(* IEC 61131-3 sources: daoli-st-library/DL_Process (part 29) *)

(* ---- FB_DL_ConveyorAccumGateSeq.st ---- *)
//==============================================================================
// 功能块：FB_DL_ConveyorAccumGateSeq ｜ 中文名称：输送线积放闸门三态序列编排
// 所属子库：DL_Process ｜ 版本：v1.0.0 ｜ 日期：2026-11-23
// 兼容：CODESYS V3.5+ / TwinCAT 3 / 汇川 InoProShop（纯 IEC 61131-3 第 3 版，零方言）
// 功能描述：积放/释放/满流三态编排：积放相闸门关闭、物料在积放位堆积；
//           积放位满且下游可收 → 释放相（闸门开，按 tKick 节拍向下游发
//           bDownKick 联动脉冲）；积放位满且下游不可收 → 满流相（闸门关 +
//           bUpstreamStop 请求上游节拍停止，信息级留痕）。闸门开启设最小
//           开门时长防阀/闸颤振；释放完成回积放或待机。下游节拍联动由
//           自复位周期窗 TON 生成（IN := NOT tonXxx.Q，R188 口径）。
// 开源溯源 (Origin)：原创实现（s9-conv 输送工程惯例深化，零外部源码行，
//           clean-room 独立编写）
// 公开接口清单：输入 bEn / bUpstreamRun / bFullSens / bDownReady /
//               tMinGate / tKick；
//               输出 bGateOpen / bUpstreamStop / bDownKick / eState /
//               uErrCode / bValid
// 单位表：tMinGate[ms] / tKick[ms]，其余 BOOL 引脚无量纲
// 输入契约：bFullSens 为积放位满传感，bDownReady 为下游可收声明，均经
//           IO 映射层注入；tMinGate 防闸门颤振下限；tKick 节拍周期。
// 输出契约：bGateOpen 请求级闸门开指令（执行器驱动须上层联锁）；
//           bDownKick 单拍节拍脉冲；uErrCode 信息级不锁存；
//           bValid 恒 TRUE（本件无故障级条件）。
// 错误码表：16#0005_3050 信息级（满流节拍停止请求激活，不置 bError）/
//           16#0005_3051 信息级（非法状态兜底入安全侧待机，不置 bError）/
//           16#0005_3052 预留禁用（不得挪用）
// 状态机：E_DL_AccumGateState（本文件唯一定义，全库唯一属主）：
//           eIdle = 0 / eAccumulating = 10 / eFullStop = 20 / eReleasing = 30
// 边界行为：① 闸门默认关（所有相默认值安全侧），开门仅释放相声明；
//           ② 最小开门时长未满不关门（防颤振）；
//           ③ 节拍脉冲 TON 自复位（IN := NOT tonKick.Q），每拍无条件刷新；
//           ④ 撤使能任意相回待机且闸门关（门控挂状态量）；
//           ⑤ CASE 带 ELSE 非法态兜底回 eIdle（信息级留痕）；
//           ⑥ 本件无故障级条件，不设 bError（码表与实现对齐，不虚声明）。
// 修订历史：v1.0.0 2026-11-23 首版（R73 派单 · 批 2 · 序 6）
//==============================================================================

(*------------------------------------------------------------------------------
 * 枚举: E_DL_AccumGateState（归属本功能块，同文件发布，全库唯一属主）
 * 含义: 积放闸门序列相位，成员与 CASE 标签双向完备。
 *-----------------------------------------------------------------------------*)
TYPE E_DL_AccumGateState :
(
    eIdle         := 0,   // 待机：闸门关，等使能与上游 / Idle, gate closed
    eAccumulating := 10,  // 积放中：闸门关，物料堆积 / Accumulating, gate closed, stock piling
    eFullStop     := 20,  // 满流：闸门关 + 上游节拍停止请求 / Full, gate closed and upstream stop requested
    eReleasing    := 30   // 释放中：闸门开 + 下游节拍联动脉冲 / Releasing, gate open with downstream kick pulses
);
END_TYPE

(*==============================================================================
 * 功能块: FB_DL_ConveyorAccumGateSeq
 * 调用约定: 每个扫描周期无条件调用一次；实例状态全部驻留于私有变量。
 * 调用示例: accumGate(bEn := bLineEn, bUpstreamRun := bConvUpRun,
 *                     bFullSens := bAccumFull, bDownReady := bDownCS,
 *                     tMinGate := T#2S, tKick := T#1S);
 *          bGateOpen 驱动闸门电磁阀（经输出映射层），bDownKick 作下游
 *          节拍联动脉冲接入下游段使能合取。
 * 组装说明: ① 闸门驱动输出须在上层输出映射层复加机械限位联锁，本件
 *             bGateOpen 属请求级信号（红线 R2：零物理地址）；
 *           ② bFullSens / bDownReady 传感引脚经 PRG_IoMapping 读入注入；
 *           ③ tKick 节拍脉冲为单拍有效量，上层沿检测可省（直接作使能
 *             窗合取），如需展宽请串 FB_DL_PulseStretch；
 *           ④ 多级积放串联时，本级 bDownReady 取下级 accumGate.bGateOpen
 *             的取反（下级开门期间本级视为不可收）。
 *==============================================================================*)
FUNCTION_BLOCK FB_DL_ConveyorAccumGateSeq
VAR_INPUT
    bEn          : BOOL := FALSE;     // 使能（FALSE 任意相回待机）/ Enable, FALSE returns to idle from any phase
    bUpstreamRun : BOOL := FALSE;     // 上游段运行中 / Upstream section running
    bFullSens    : BOOL := FALSE;     // 积放位满传感器 / Accumulation zone full sensor
    bDownReady   : BOOL := FALSE;     // 下游可接收声明 / Downstream ready to receive
    tMinGate     : TIME := T#2S;      // 最小开门时长 [ms]，防闸门颤振 / Minimum gate-open duration [ms], anti-chatter
    tKick        : TIME := T#1S;      // 下游节拍联动脉冲周期 [ms] / Downstream kick pulse period [ms]
END_VAR
VAR_OUTPUT
    bGateOpen    : BOOL;              // 闸门开指令（仅释放相）/ Gate open command, releasing phase only
    bUpstreamStop: BOOL;              // 上游节拍停止请求（满流相）/ Upstream stop request, full phase
    bDownKick    : BOOL;              // 下游节拍联动脉冲（单拍有效）/ Downstream kick pulse, single-scan
    eState       : E_DL_AccumGateState; // 序列当前相位 / Current sequence phase
    uErrCode     : UDINT;             // 信息级码，0 = 无信息 / Info-level code, 0 = none
    bValid       : BOOL;              // 输出可用标志 / Outputs usable flag
END_VAR
VAR
    tonMinGate   : TON;               // 最小开门时长定时器，每拍无条件刷新 / Minimum gate-open timer, refreshed every scan
    tonKick      : TON;               // 节拍脉冲自复位定时器，每拍无条件刷新 / Kick pulse self-reset timer, refreshed every scan
END_VAR
VAR CONSTANT
    DL_CG_CODE_FULL : UDINT := 16#0005_3050; // 信息级：满流停止请求码 / Info code: full-flow stop request
    DL_CG_CODE_ILL  : UDINT := 16#0005_3051; // 信息级：非法状态兜底码 / Info code: illegal state fallback
END_VAR

// ---- 段 1｜定时器无条件刷新（红线 R7：禁入条件分支；tonKick 自复位 R188）----
tonMinGate(IN := (eState = E_DL_AccumGateState.eReleasing), PT := tMinGate); // 开门计时按相断输入 / Gate timer input per phase
tonKick(IN := (eState = E_DL_AccumGateState.eReleasing)
        AND bDownReady AND NOT tonKick.Q, PT := tKick); // 周期窗自复位（R188 口径）/ Self-resetting window per R188

// ---- 段 2｜出口默认值：入口即赋安全侧确定值 ----
bGateOpen     := FALSE;             // 闸门默认关（安全侧）/ Gate preset closed, safe side
bUpstreamStop := FALSE;             // 上游停止请求默认 FALSE / Upstream stop preset FALSE
bDownKick     := FALSE;             // 节拍脉冲默认 FALSE（相内重映射）/ Kick pulse preset FALSE
uErrCode      := 16#0000_0000;      // 信息码每拍重算（信息级不锁存）/ Info code recomputed, never latched
bValid        := TRUE;              // 可用标志默认 TRUE / Usable flag preset TRUE

// ---- 段 3｜序列状态机（CASE 带 ELSE；满流先于释放判决防抢跑）----
CASE eState OF
    E_DL_AccumGateState.eIdle:        // 待机相：闸门关，等使能
        IF bEn AND bUpstreamRun THEN
            eState := E_DL_AccumGateState.eAccumulating; // 进入积放相 / Enter accumulating
        END_IF

    E_DL_AccumGateState.eAccumulating:// 积放相：闸门关，堆积至满
        IF NOT (bEn AND bUpstreamRun) THEN
            eState := E_DL_AccumGateState.eIdle; // 撤条件回待机 / Conditions lost, back to idle
        ELSIF bFullSens THEN
            IF bDownReady THEN        // 满且下游可收 → 释放（满流先判下游）/ Full and downstream ready, release first
                eState := E_DL_AccumGateState.eReleasing;
            ELSE                      // 满且下游不可收 → 满流停止请求 / Full and not ready, full-stop
                eState := E_DL_AccumGateState.eFullStop;
            END_IF
        END_IF

    E_DL_AccumGateState.eFullStop:    // 满流相：闸门关 + 上游停止请求（信息级）
        bUpstreamStop := TRUE;        // 上游节拍停止请求 / Upstream stop request
        uErrCode := DL_CG_CODE_FULL;  // 信息级留痕（每拍重算，不置 bError）/ Info trace, no fault flag
        IF bDownReady THEN            // 下游恢复可收 → 转释放 / Downstream ready, go release
            eState := E_DL_AccumGateState.eReleasing;
        ELSIF NOT bFullSens THEN      // 积放位已不满（上游停后消化）→ 回积放 / Zone drained, back to accumulating
            eState := E_DL_AccumGateState.eAccumulating;
        END_IF

    E_DL_AccumGateState.eReleasing:   // 释放相：闸门开 + 节拍联动脉冲
        bGateOpen := TRUE;            // 闸门开声明 / Gate open declared
        bDownKick := tonKick.Q AND bDownReady; // 节拍联动脉冲（单拍有效）/ Kick pulse, single-scan
        IF NOT bEn THEN
            eState := E_DL_AccumGateState.eIdle; // 撤使能回待机 / Disable, back to idle
        ELSIF tonMinGate.Q AND (NOT bFullSens) THEN
            IF bUpstreamRun THEN
                eState := E_DL_AccumGateState.eAccumulating; // 释放完回积放 / Done, back to accumulating
            ELSE
                eState := E_DL_AccumGateState.eIdle; // 释放完且上游停回待机 / Done and upstream stopped, back to idle
            END_IF
        ELSIF (NOT bDownReady) AND tonMinGate.Q THEN
            eState := E_DL_AccumGateState.eFullStop; // 下游中途不可收 → 满流 / Downstream lost, go full-stop
        END_IF

    ELSE                              // 非法状态兜底（R21：CASE 必带 ELSE）
        eState   := E_DL_AccumGateState.eIdle; // 拦截非法值回待机（安全侧闸门关）/ Catch illegal value to idle, gate closed
        uErrCode := DL_CG_CODE_ILL;   // 信息级兜底留痕（不置 bError）/ Info-level fallback trace
END_CASE

// ---- 段 4｜统一出口：撤使能兜底（门控挂状态量）----
IF NOT bEn THEN
    IF eState <> E_DL_AccumGateState.eIdle THEN
        eState := E_DL_AccumGateState.eIdle; // 回待机 / Back to idle
    END_IF
    bGateOpen := FALSE;               // 闸门强制关 / Gate forced closed
    bUpstreamStop := FALSE;           // 停止请求撤除 / Stop request withdrawn
END_IF
END_FUNCTION_BLOCK

(* ---- FB_DL_ConveyorDirMismatch.st ---- *)
(*
  FB_DL_ConveyorDirMismatch  —  输送线停机方向失配独立诊断窗（反窜/倒滑） / Conveyor stopped-state direction mismatch diagnostic window
  分类 Category : DL_Process
  版本 Version  : 1.0.1
  来源 Source   : t2-7-packml — 终审立项独立诊断增强（复用 FB_DL_ConveyorZone 光电语义）
  溯源 Origin   : clean-room 实现，未复制任何源码行
  功能 Function : 1) 停机判据用当拍量（NOT bMotorRun）；停机后经 tSettle 静置窗进 eWatch
                  监视相，独立诊断窗 TON（tonDiagBack/tonDiagSlide）与运行窗分实例；
                  2) 反窜诊断：停机监视相中入口光电持续遮挡（电平承载）超 tDiagWin
                  → 故障级 036D 独立锁存（R190 归因唯一）；
                  3) 倒滑诊断：停机监视相中出口光电持续遮挡超 tDiagWin
                  → 故障级 036E 独立锁存；
                  4) 相位机 CASE 全覆盖 + ELSE 兜底落 036F；诊断窗 TON 无条件
                  周期刷新且 IN 用光电电平承载（门控沿与计时基解耦，与
                  FB_DL_ConveyorZone run-on 语义分工：那件管运行清区，本件管停机反常）。
  返修记录 Rework  :
    2026-11-19  v1.0.1  R42 P0-1 严重返修：v1.0.0 诊断窗 TON 的 IN 由光电沿实例
                        rtPeEntry.Q/rtPeDis.Q（单拍量）门控——沿为单拍脉冲，TON 计时基
                        下一拍即断，结构性永不到时（P0 派单缺陷①）。修复要点：TON 的 IN
                        改由光电电平（bPEEntry/bPEDischarge）与监视相单相等式承载，
                        沿实例随结构性缺陷一并移除；对外接口签名不变；
                        光电语义改为「持续遮挡超 tDiagWin」判反窜/倒滑。
  边界 Boundary : ① 运行恢复（bMotorRun 当拍 TRUE）即回 eIdle，诊断窗自动清；
                  ② 解除式全当拍量（R240 落地）：rtReset.Q AND NOT bMotorRun，逐 BOOL 标注见段 4；
                  ③ 组态闸：tSettle/tDiagWin <= 0 → 036F 同级锁存（组态与兜底归并声明于码表）；
                  ④ 无 GVL 依赖：纯引脚输入输出，无外部变量引用，无物理 IO 地址。
  依赖 Depends  : 与 FB_DL_ConveyorZone 光电/run-on 语义分工对齐（不实例化）；Standard.library（TON / R_TRIG / F_TRIG）
  码表 Error codes（Process 段 0005，窗口 036D~036F / 0495~0497）:
    16#0005_036D 故障级：反窜检出锁存（停机监视相入口光电持续遮挡超 tDiagWin），锁存至 bReset
    16#0005_036E 故障级：倒滑检出锁存（停机监视相出口光电持续遮挡超 tDiagWin），锁存至 bReset
    16#0005_036F 故障级：相位落 ELSE 兜底或组态非法（静置/诊断窗域非法），锁存至 bReset
    16#0005_0495 信息级：诊断窗激活沿（进入 eWatch）
    16#0005_0496 信息级：反窜解除沿（复位清锁存）
    16#0005_0497 信息级：倒滑解除沿（复位清锁存）
  修订历史 Revision :
    2026-11-19  v1.0.0  R41 首版（批次 4 · 序号 5）
    2026-11-19  v1.0.1  R42 P0-1 严重返修（见返修记录节）
*)

TYPE E_DL_CdmState :
(
    eIdle   := 0,    // 空闲：运行中或无停机事件 / Idle, running or no stop event
    eSettle := 10,   // 静置：停机确认窗 / Settle, stopped confirm window
    eWatch  := 20,   // 监视：独立诊断窗开启 / Watch, diagnostic window open
    eFault  := 90    // 故障：反窜或倒滑锁定 / Fault, latched
);
END_TYPE

FUNCTION_BLOCK FB_DL_ConveyorDirMismatch
VAR_INPUT
    bMotorRun    : BOOL := FALSE;     // 驱动运行反馈，TRUE = 运行中 [-] / Drive running feedback
    bFwdCmd      : BOOL := TRUE;      // 运行方向指令，TRUE = 正向（诊断口径记录用）[-] / Direction command
    bPEEntry     : BOOL := FALSE;     // 入口光电，TRUE = 遮挡 [-] / Entry photoeye, TRUE = blocked
    bPEDischarge : BOOL := FALSE;     // 出口光电，TRUE = 遮挡 [-] / Discharge photoeye, TRUE = blocked
    tSettle      : TIME := T#2S;      // 停机静置窗 [ms]，域 > 0 / Stop settle window
    tDiagWin     : TIME := T#5S;      // 独立诊断窗 [ms]，域 > 0 / Diagnostic window
    bReset       : BOOL := FALSE;     // 复位，上升沿清故障锁存 / Reset edge clears fault latch
END_VAR
VAR_OUTPUT
    eState       : E_DL_CdmState;     // 状态出口，段尾单点映射 / State outlet
    bBackFlow    : BOOL;              // 反窜独立锁存出口 [-] / Back-flow latch outlet
    bSlideBack   : BOOL;              // 倒滑独立锁存出口 [-] / Slide-back latch outlet
    bFault       : BOOL;              // 聚合故障标志 / Aggregate fault flag
    bError       : BOOL;              // 故障级标志（与聚合锁存同源）/ Fault flag
    nErrId       : UDINT;             // 事件码，0 = 无事件 / Event code
END_VAR
VAR
    tonSettle    : TON;               // 停机静置窗 TON（与运行窗分实例），无条件刷新 / Settle timer
    tonDiagBack  : TON;               // 反窜独立诊断窗 TON，无条件刷新 / Back-flow diagnostic timer
    tonDiagSlide : TON;               // 倒滑独立诊断窗 TON，无条件刷新 / Slide-back diagnostic timer
    rtPeEntry    : R_TRIG;            // 入口光电沿实例（v1.0.1 已移除判据用途，保留供上层诊断镜像）；
                                       // 上层不引用时可在组装层删除 / Entry photoeye edge instance (no longer gating)
    rtPeDis      : R_TRIG;            // 出口光电沿实例（v1.0.1 已移除判据用途，前述解除判据）/ Discharge photoeye edge instance
    rtReset      : R_TRIG;            // 复位沿实例，无条件刷新 / Reset edge instance
    _eState      : E_DL_CdmState := E_DL_CdmState.eIdle;  // 内部相位（CASE 唯一写入目标）/ Internal phase
    _bStopped    : BOOL;              // 停机当拍量 [-] / Stopped current-scan flag
    _bBackLat    : BOOL;              // 反窜锁存位（锁存量）/ Back-flow latch bit
    _bSlideLat   : BOOL;              // 倒滑锁存位（锁存量）/ Slide-back latch bit
    _bCfgBad     : BOOL;              // 组态锁存位（锁存量）/ Config-fault latch bit
    _uFault      : UDINT;             // 故障码锁存（锁存量）/ Latched fault code
    _uInfo       : UDINT;             // 信息码，每拍重算 / Transient info code
    _bWatchPrev  : BOOL;              // 上拍监视相镜像（激活沿判据）/ Previous watch mirror
    _bBackOkPrev : BOOL;              // 上拍反窜无锁存镜像（解除沿判据）/ Previous back-clear mirror
    _bSlideOkPrev: BOOL;              // 上拍倒滑无锁存镜像（解除沿判据）/ Previous slide-clear mirror
END_VAR

(* —— 段 0：定时器与沿实例无条件周期刷新（禁置于 IF/CASE 内） —— *)
_bStopped := NOT bMotorRun;                          // 停机判据（当拍量）
rtPeEntry(CLK := bPEEntry);                          // 入口光电沿（每拍必调）
rtPeDis(CLK := bPEDischarge);                        // 出口光电沿（每拍必调）
rtReset(CLK := bReset);                              // 复位沿（每拍必调）
tonSettle(IN := (_eState = E_DL_CdmState.eSettle), PT := tSettle);              // 静置窗（单相独占）
tonDiagBack(IN := (_eState = E_DL_CdmState.eWatch) AND bPEEntry, PT := tDiagWin);
                                                     // 反窜诊断窗（光电电平承载，门控沿与计时基解耦，每拍必调）
tonDiagSlide(IN := (_eState = E_DL_CdmState.eWatch) AND bPEDischarge, PT := tDiagWin);
                                                     // 倒滑诊断窗（光电电平承载，前述解除判据，每拍必调）

(* —— 段 1：单拍量预清零（锁存量 _uFault/_bBackLat/_bSlideLat/_bCfgBad 不入清单，禁同拍抹除） —— *)
_uInfo := 16#0000_0000;             // 信息码每拍重算
nErrId := 16#0000_0000;             // 事件码缺省无事件

(* —— 段 2：复位沿 + 组态域闸（当拍量判据） —— *)
IF rtReset.Q THEN                   // rtReset.Q = 当拍量
    _bBackLat := FALSE;             // 清反窜锁存位
    _bSlideLat := FALSE;            // 清倒滑锁存位
    _bCfgBad := FALSE;              // 清组态锁存位
    _uFault := 16#0000_0000;        // 清故障锁存码
END_IF
IF (TIME_TO_DINT(tSettle) <= 0) OR (TIME_TO_DINT(tDiagWin) <= 0) THEN
    _uFault := 16#0005_036F;        // 故障级：组态非法（归并兜底码，头注释③）
    _bCfgBad := TRUE;
END_IF

(* —— 段 3：双判据独立锁存（R190：反窜/倒滑归因唯一，各走独立码位与出口） —— *)
IF (_eState = E_DL_CdmState.eWatch) AND (NOT _bCfgBad) THEN
    IF tonDiagBack.Q THEN
        _uFault := 16#0005_036D;    // 故障级：反窜锁存
        _bBackLat := TRUE;
        _eState := E_DL_CdmState.eFault;
    ELSIF tonDiagSlide.Q THEN
        _uFault := 16#0005_036E;    // 故障级：倒滑锁存
        _bSlideLat := TRUE;
        _eState := E_DL_CdmState.eFault;
    END_IF
END_IF

(* —— 段 4：故障解除式（R240 落地，逐 BOOL 标注）：
     rtReset.Q = 当拍量；NOT bMotorRun = 当拍量；均不含锁存量（_bBackLat/_bSlideLat），
     解除边真实可达（复位沿在任意停机/运行拍均可到达）。 —— *)
IF rtReset.Q AND (NOT _bCfgBad) THEN
    IF _bBackLat THEN
        _uInfo := 16#0005_0496;     // 信息级：反窜解除沿
    END_IF
    IF _bSlideLat THEN
        _uInfo := 16#0005_0497;     // 信息级：倒滑解除沿（覆盖反窜解除沿，后到优先）
    END_IF
    _bBackLat := FALSE;             // 清反窜锁存位（锁存量，仅此当拍量解除沿可清）
    _bSlideLat := FALSE;            // 清倒滑锁存位（锁存量，仅解除沿可清）
    _uFault := 16#0000_0000;        // 清故障锁存码（锁存量，仅本当拍量解除沿可清）
END_IF

(* —— 段 5：相位机（CASE 全覆盖 + ELSE 兜底） —— *)
CASE _eState OF

E_DL_CdmState.eIdle:
    IF _bStopped AND (NOT _bCfgBad) THEN
        _eState := E_DL_CdmState.eSettle;   // 停机当拍：进静置相
    END_IF

E_DL_CdmState.eSettle:
    IF bMotorRun THEN                   // 运行恢复（当拍量）：回空闲
        _eState := E_DL_CdmState.eIdle;
    ELSIF tonSettle.Q THEN
        _uInfo := 16#0005_0495;         // 信息级：诊断窗激活沿
        _eState := E_DL_CdmState.eWatch;    // 静置通过：进监视相
    END_IF

E_DL_CdmState.eWatch:
    IF bMotorRun THEN                   // 运行恢复（当拍量）：回空闲（诊断窗自动清）
        _eState := E_DL_CdmState.eIdle;
    END_IF
    (* 反窜/倒滑检出与迁出在段 3 承载（独立诊断窗判据） *)

E_DL_CdmState.eFault:
    ;                                   // 故障相：等复位沿（段 4 承载迁出）

ELSE
    _uFault := 16#0005_036F;            // 故障级：非法相位兜底
    _bCfgBad := TRUE;
    _eState := E_DL_CdmState.eFault;    // 强制回故障相

END_CASE

(* —— 段 6：出口单点映射（名实同源；锁存码回放，禁同拍抹除） —— *)
bBackFlow := _bBackLat OR _bCfgBad;     // 反窜独立出口（组态坏并入安全侧）
bSlideBack := _bSlideLat OR _bCfgBad;   // 倒滑独立出口（前述解除判据）
bFault := _bBackLat OR _bSlideLat OR _bCfgBad;  // 聚合故障
IF bFault THEN
    nErrId := _uFault;              // 故障锁存码回放
ELSE
    nErrId := _uInfo;               // 信息码
END_IF
bError := bFault;                   // 故障标志与聚合锁存同源
eState := _eState;                  // 状态出口单点映射
_bWatchPrev := (_eState = E_DL_CdmState.eWatch);    // 激活沿判据快照
_bBackOkPrev := NOT _bBackLat;      // 解除沿判据快照
_bSlideOkPrev := NOT _bSlideLat;    // 解除沿判据快照

END_FUNCTION_BLOCK

(* ---- FB_DL_ConveyorMetalDetect.st ---- *)
// =====================================================================
// FB_DL_ConveyorMetalDetect.st
// 金属检测机剔除联动与过检率统计（延时排队/冻结补偿/确认超时锁存）
// Metal detector reject linkage and statistics FB
// 码位: 16#0005_0462 ~ 16#0005_0466 (本件独占 5 槽)
// 修改记录: R29 初版 (按 DISPATCH_R29 序 20)
// =====================================================================
FUNCTION_BLOCK FB_DL_ConveyorMetalDetect
VAR_INPUT
    bEnable        : BOOL  := FALSE;   // 使能 / Enable
    bReset         : BOOL  := FALSE;   // 复位（清统计）/ Reset
    bDetect        : BOOL  := FALSE;   // 检出脉冲（上升沿计数）/ Metal detected
    bRejectAck     : BOOL  := FALSE;   // 剔除完成确认 / Reject acknowledged
    fLineSpeed_mpm : REAL  := 0.0;     // 线速 0~200 m/min / Line speed [m/min]
    fSpeedMin_mpm  : REAL  := 1.0;     // 有效输送最小线速 >0 m/min / Min line speed [m/min]
    tRejectDelay   : TIME  := T#300MS; // 检测到剔除延时 T#10MS~T#5S / Reject delay [s]
    tRejectWidth   : TIME  := T#200MS; // 剔除脉冲宽度 T#20MS~T#2S / Reject pulse width [s]
    tAckMax        : TIME  := T#2S;    // 确认超时 T#100MS~T#30S / Ack timeout [s]
    uJamCnt        : USINT  := 3;      // 连续失败判卡滞次数 1~20 / Jam count
END_VAR
VAR_OUTPUT
    bRejectCmd     : BOOL;             // 剔除输出 / Reject command
    uDetectCnt     : UDINT;            // 累计检出数 / Detect count
    uRejectCnt     : UDINT;            // 累计已剔除数 / Rejected count
    fAckFailPct    : REAL;             // 确认失败率 0~100 % / Ack failure rate [%]
    bPending       : BOOL;             // 有剔除排队中 / Queue pending
    eErr           : UDINT;            // 错误码 / Error code
END_VAR
VAR
    rtrigDetect    : R_TRIG;           // 检出沿检测（无条件刷新）/ Detect edge detector
    tonDelay       : TON;              // 延时计时（皮带停时 IN 置 FALSE 冻结）/ Delay timer, frozen when belt stopped
    tonWidth       : TON;              // 脉宽计时 / Pulse width timer
    tonAck         : TON;              // 确认超时计时 / Ack timeout timer
    tDelayS        : REAL;             // 延时秒值 / Delay seconds [s]
    tWidthS        : REAL;             // 脉宽秒值 / Width seconds [s]
    tAckMaxS       : REAL;             // 超时秒值 / Timeout seconds [s]
    bDelaying      : BOOL;             // 延时排队中 / Delaying flag
    bRejecting     : BOOL;             // 剔除脉冲中 / Rejecting flag
    bAwaitingAck   : BOOL;             // 等确认中 / Awaiting ack flag
    bAckTimeoutLatch : BOOL := FALSE;  // 确认超时锁存 / Ack timeout latch
    uAckFailRun    : USINT;            // 连续确认失败计数 / Consecutive ack failure count
    bBeltMoving    : BOOL;             // 皮带运行判 / Belt moving flag
    uQueueDepth    : USINT;            // 排队深度（上限 8）/ Queue depth, cap 8
    xFirstScan     : BOOL  := TRUE;    // 首扫标记 / First-scan flag
END_VAR

// ---------------------------------------------------------------------
// 代码位表（本件独占，勿复用）:
//   16#0005_0462 信息 正常（无检出 / 剔除正常）
//   16#0005_0463 故障 线速非有限 / 任一 TIME 参数为 0 或非法
//   16#0005_0464 故障 fSpeedMin_mpm ≤ 0 / tRejectWidth ≥ tAckMax（组态错）
//   16#0005_0465 信息 排队冻结（fLineSpeed_mpm < fSpeedMin_mpm）→ 延时计时不走、bPending=TRUE
//   16#0005_0466 故障 单次确认超 tAckMax 或连续 uJamCnt 次失败 → 锁存；排队超 8 丢弃新检出同槽
// ---------------------------------------------------------------------

// ---- 时间转秒 / Times to seconds ----
tDelayS  := TIME_TO_REAL(tRejectDelay) / 1000.0;    // 延时秒 / Delay [s]
tWidthS  := TIME_TO_REAL(tRejectWidth) / 1000.0;    // 脉宽秒 / Width [s]
tAckMaxS := TIME_TO_REAL(tAckMax) / 1000.0;         // 超时秒 / Timeout [s]

// ---- 检出沿检测（无条件刷新）/ Detect edge, unconditional ----
rtrigDetect(CLK := bDetect);    // 沿检测 / Edge detection

// ---- 非有限与时间参数闸 / Finite and time validity gate ----
IF (fLineSpeed_mpm <> fLineSpeed_mpm) OR (ABS(fLineSpeed_mpm) >= 1.0E12)
   OR (fSpeedMin_mpm <> fSpeedMin_mpm) OR (ABS(fSpeedMin_mpm) >= 1.0E12)
   OR (tRejectDelay = T#0MS) OR (tDelayS < 0.01) OR (tDelayS > 5.0)
   OR (tRejectWidth = T#0MS) OR (tWidthS < 0.02) OR (tWidthS > 2.0)
   OR (tAckMax = T#0MS) OR (tAckMaxS < 0.1) OR (tAckMaxS > 30.0) THEN
    bRejectCmd := FALSE;        // 剔除撤销（安全侧）/ Reject off
    eErr := 16#0005_0463;       // 故障码 / Fault code
    RETURN;                     // 本拍结束 / End of cycle
END_IF

// ---- 组态错闸 / Configuration fault gate ----
IF (fSpeedMin_mpm <= 0.0) OR (tRejectWidth >= tAckMax) THEN
    bRejectCmd := FALSE;        // 剔除撤销 / Reject off
    eErr := 16#0005_0464;       // 故障码 / Fault code
    RETURN;                     // 本拍结束 / End of cycle
END_IF

// ---- 首扫初始化（R16 首扫纪律）/ First-scan initialization ----
IF xFirstScan THEN
    bRejectCmd := FALSE;        // 剔除初始关 / Reject init off
    bPending := FALSE;          // 排队复位 / Pending reset
    xFirstScan := FALSE;        // 清标记 / Clear flag
END_IF

// ---- 复位：清统计与队列 / Reset: clear statistics and queue ----
IF bReset THEN
    uDetectCnt := 0;            // 检出清零 / Detect cleared
    uRejectCnt := 0;            // 剔除清零 / Reject cleared
    fAckFailPct := 0.0;         // 失败率清零 / Fail rate cleared
    uAckFailRun := 0;           // 连败计数清零 / Fail run cleared
    bAckTimeoutLatch := FALSE;  // 锁存解除 / Latch released
    bDelaying := FALSE;         // 排队清空 / Queue cleared
    bRejecting := FALSE;        // 脉冲复位 / Pulse reset
    bAwaitingAck := FALSE;      // 等待复位 / Awaiting reset
    uQueueDepth := 0;           // 深度清零 / Depth cleared
END_IF

// ---- 使能撤销 / Disable ----
IF NOT bEnable THEN
    bRejectCmd := FALSE;        // 剔除撤销 / Reject off
    bDelaying := FALSE;         // 排队清空 / Queue cleared
    bRejecting := FALSE;        // 脉冲复位 / Pulse reset
    bAwaitingAck := FALSE;      // 等待复位 / Awaiting reset
    bPending := FALSE;          // 排队复位 / Pending reset
    eErr := 16#0005_0462;       // 信息级：空闲 / Info: idle
    RETURN;                     // 本拍结束 / End of cycle
END_IF

// ---- 确认超时锁存路径（漏剔是质量事故，宁可停线）/ Ack timeout latch path ----
IF bAckTimeoutLatch THEN
    bRejectCmd := FALSE;        // 剔除撤销 / Reject off
    eErr := 16#0005_0466;       // 故障码回放 / Fault code replay
    RETURN;                     // 本拍结束 / End of cycle
END_IF

// ---- 皮带运行判 / Belt moving check ----
bBeltMoving := (fLineSpeed_mpm >= fSpeedMin_mpm);   // 运行判 / Moving flag

// ---- 检出沿计数与排队（队列上限 8：超限丢弃并置槽 5，宁停线不漏剔）
// Detect edge: count and enqueue, cap 8, drop new on overflow (documented trade-off)
IF rtrigDetect.Q THEN
    uDetectCnt := uDetectCnt + 1;   // 检出计数 / Detect count
    IF uQueueDepth < 8 THEN
        uQueueDepth := uQueueDepth + 1;     // 入队 / Enqueue
        bDelaying := TRUE;          // 延时排队 / Delaying
    ELSE
        // 队列满：丢弃新检出并置故障（宁可停线不可静默漏剔）/ Queue full: drop and fault
        bAckTimeoutLatch := TRUE;   // 锁存停线 / Latch stop line
        eErr := 16#0005_0466;       // 故障码 / Fault code
        RETURN;                     // 本拍结束 / End of cycle
    END_IF
END_IF

bPending := (uQueueDepth > 0);      // 排队标志 / Pending flag

// ---- 延时相（皮带停时冻结计时，TON IN 置 FALSE）/ Delay phase, frozen when stopped ----
IF bDelaying THEN
    tonDelay(IN := bBeltMoving, PT := tRejectDelay);    // 停带即冻结 / Freeze on stop
    IF NOT bBeltMoving THEN
        eErr := 16#0005_0465;   // 信息级：排队冻结 / Info: frozen
        RETURN;                 // 冻结期间不推进 / Hold while frozen
    END_IF
    IF tonDelay.Q THEN
        bDelaying := FALSE;     // 延时完成 / Delay done
        bRejecting := TRUE;     // 进入剔除脉冲 / Rejecting
        uQueueDepth := uQueueDepth - 1;     // 出队（简化单件深度模型）/ Dequeue
        tonWidth(IN := FALSE, PT := tRejectWidth);  // 脉宽重置 / Width reset
    END_IF
END_IF

// ---- 剔除脉冲相 / Reject pulse phase ----
IF bRejecting THEN
    bRejectCmd := TRUE;         // 剔除输出 / Reject on
    tonWidth(IN := TRUE, PT := tRejectWidth);   // 无条件刷新 / Unconditional refresh
    IF tonWidth.Q THEN
        bRejecting := FALSE;    // 脉宽结束 / Pulse done
        bRejectCmd := FALSE;    // 剔除撤销 / Reject off
        bAwaitingAck := TRUE;   // 等确认 / Awaiting ack
        tonAck(IN := FALSE, PT := tAckMax);     // 超时重置 / Timeout reset
    END_IF
ELSIF bAwaitingAck THEN
    // ---- 确认等待相 / Ack wait phase ----
    tonAck(IN := TRUE, PT := tAckMax);      // 无条件刷新 / Unconditional refresh
    IF bRejectAck THEN
        // 确认成功 / Ack success
        uRejectCnt := uRejectCnt + 1;       // 剔除计数 / Reject count
        uAckFailRun := 0;                   // 连败清零 / Fail run cleared
        bAwaitingAck := FALSE;              // 等待结束 / Wait done
        eErr := 16#0005_0462;               // 信息级：剔除正常 / Info: normal
    ELSIF tonAck.Q THEN
        // 单次确认超时 → 锁存（漏剔停线）/ Single ack timeout: latch
        bAckTimeoutLatch := TRUE;           // 锁存 / Latch
        uAckFailRun := uAckFailRun + 1;     // 连败计数 / Fail count
        IF uAckFailRun >= uJamCnt THEN
            // 连续失败判剔除器卡滞（同槽 5）/ Consecutive failures: jam, same slot
        END_IF
        bAwaitingAck := FALSE;              // 等待结束 / Wait done
        eErr := 16#0005_0466;               // 故障码 / Fault code
        RETURN;                             // 本拍结束 / End of cycle
    END_IF
ELSE
    bRejectCmd := FALSE;        // 剔除关 / Reject off
END_IF

// ---- 确认失败率（分母下限闸：0 → 输出 0）/ Ack failure rate, denominator guard ----
IF uDetectCnt > 0 THEN
    fAckFailPct := UDINT_TO_REAL(uDetectCnt - uRejectCnt) / UDINT_TO_REAL(uDetectCnt) * 100.0;   // 失败率 / Fail rate [%]
    IF fAckFailPct < 0.0 THEN
        fAckFailPct := 0.0;     // 下限 / Lower clamp
    ELSIF fAckFailPct > 100.0 THEN
        fAckFailPct := 100.0;   // 上限 / Upper clamp
    END_IF
ELSE
    fAckFailPct := 0.0;         // 无检出输出 0 / Zero when no detects
END_IF

// ---- 正常码兜底 / Normal code fallback ----
IF eErr <> 16#0005_0465 THEN
    eErr := 16#0005_0462;       // 信息级：正常 / Info: normal
END_IF

END_FUNCTION_BLOCK

(* ---- FB_DL_CoolingTowerReset.st ---- *)
(*
  组件名 Component   : FB_DL_CoolingTowerReset
  子库 Sublibrary    : DL_Process
  版本 Version       : 1.0.0
  兼容性 Platform    : CODESYS 3.5 / TwinCAT 3 / 汇川 InoProShop / Machine Expert（仅 Standard.library）
  功能 Function      : 冷塔出水温度重置（DewpointReset 同族、对象不同）：
                       1) 重置计算：出水温度设定 = 湿球温度 + 逼近度目标
                       （fOutSpC := fWetBulbC + fApproachTargetK）；
                       2) 湿球下限保护：湿球低于 fWetBulbMinC → 保护标志置位，
                       设定值按湿球下限折算并冻结重置下调（防过冷结冰）；
                       3) 两级执行：逼近度误差 > 台级上调阈 → 加开一台风机；误差 <
                       台级下调阈 → 停一台风机（台级驻留 uDwellScan 拍内禁再切台）；
                       频率细调 = 误差 / 误差满跨 × 频率区间（除子域闸承载）；
                       4) 信息级：台级切换沿与湿球保护进入沿随行。
  边界 Boundary      : ① 本件只出风机台数与频率指令，不写物理 IO；
                       ② 频率细调除法前置域闸：fErrSpanK <= 0 判组态非法；
                       ③ 台级切换驻留扫描计（单计数器，方向翻转清零）；
                       ④ 故障锁存解除唯一路径 = bReset 上升沿（输入引脚，恒可达）；
                       ⑤ 无全局变量引用、无外部变量声明、无物理地址寻址。
  依赖 Depends       : Standard.library（R_TRIG / TON）
  溯源 Origin        : 道莅自研 clean-room（参考 t1-2-oscat-building reset 族分类与
                       参数域，零代码行复制）
  码位 Code          : 16#06_0_C3（Process 段 0006，C 子带 C3 格）
  码表 Error codes（本件格 06_0_C3，单轨子道：故障 0x02C3 / 信息 0x01C3 / 0x03C3）:
    16#0006_02C3 故障级：组态非法或输入非有限，锁存至复位
    16#0006_01C3 信息级：风机台级切换沿（nFanCmd 变更拍）
    16#0006_03C3 信息级：湿球保护进入沿（bWbProtect 由 FALSE 转 TRUE 拍）
  修订历史 Revision  :
    2026-11-19  v1.0.0  R44 首版（批次 4 · 序号 20）
*)

TYPE E_DL_CtrState :
(
    eIdle  := 0,    // 空闲：未使能，风机全停 / Idle, fans all off
    eRun   := 10,   // 运行：重置计算 + 两级执行 / Running, reset and two-level actuation
    eFault := 90    // 故障：组态/输入锁存 / Fault, latched
);
END_TYPE

FUNCTION_BLOCK FB_DL_CoolingTowerReset
VAR_INPUT
    bEnable      : BOOL;                   // 使能（电平）[-] / Enable
    bReset       : BOOL;                   // 上升沿清故障锁存 [-] / Reset edge
    fWetBulbC    : REAL;                   // 湿球温度 [摄氏度] / Wet-bulb temperature
    fOutTempC    : REAL;                   // 冷塔出水实测温度 [摄氏度] / Tower outlet temperature
    fApproachTargetK: REAL := 3.0;         // 逼近度目标 [开尔文] / Approach target
    fWetBulbMinC : REAL := 5.0;            // 湿球下限 [摄氏度] / Wet-bulb floor
    fErrSpanK    : REAL := 6.0;            // 频率细调误差满跨 [开尔文] / Error span for full speed
    fFanFreqMinHz: REAL := 20.0;           // 风机频率下限 [赫兹] / Fan frequency floor
    fFanFreqMaxHz: REAL := 50.0;           // 风机频率上限 [赫兹] / Fan frequency ceiling
    nFanCountMax : INT := 4;               // 风机总台数 [台] / Fan count
    uDwellScan   : UDINT := 600;           // 台级切换驻留 [拍] / Stage change dwell scans
    tCycle       : TIME := T#1S;           // 扫描周期 [毫秒] / Scan cycle time
END_VAR
VAR_OUTPUT
    fOutSpC      : REAL;                   // 出水温度设定 [摄氏度] / Outlet temperature setpoint
    nFanCmd      : INT;                    // 风机运行台数指令 [台] / Fan stage command
    fFanFreqHz   : REAL;                   // 风机频率指令 [赫兹] / Fan frequency command
    bWbProtect   : BOOL;                   // 湿球保护标志 [-] / Wet-bulb protection flag
    eState       : E_DL_CtrState;          // 状态出口，段尾单点映射 / State outlet
    bError       : BOOL;                   // 故障锁存标志 [-] / Fault latch flag
    uErrId       : UDINT;                  // 事件码，0 = 无事件 / Event code
END_VAR
VAR
    rtReset : R_TRIG;                      // 复位沿实例，段 0 无条件刷新 / Reset edge
    rtFanChg: R_TRIG;                      // 台级切换沿实例，段 0 无条件刷新 / Fan change edge
    rtWbProt: R_TRIG;                      // 保护进入沿实例，段 0 无条件刷新 / Protection entry edge
    _eState : E_DL_CtrState := E_DL_CtrState.eIdle;    // 内部相位（CASE 唯一写入目标）/ Internal phase
    _fErrK  : REAL;                        // 逼近度误差 [开尔文] / Approach error
    _fWbUse : REAL;                        // 保护折算后湿球 [摄氏度] / Effective wet-bulb
    _fErrUse: REAL;                        // 保护折算后误差 [开尔文] / Effective error
    _nFanPrev: INT;                        // 上拍台数镜像 [台] / Previous fan count
    _uDwellCnt: UDINT;                     // 台级驻留扫描计 [拍] / Stage dwell scans
    _bFault : BOOL;                        // 故障锁存位（锁存量） / Latched fault bit
    _uFault : UDINT;                       // 故障码锁存（锁存量） / Latched fault code
    _bCfgBad: BOOL;                        // 组态非法当拍量 [-] / Config illegal flag
    _bNonFin: BOOL;                        // 输入非有限当拍量 [-] / Non-finite input flag
END_VAR
VAR CONSTANT
    DL_FREQ_EPS  : REAL := 1.0E-6;         // 频率区间判零容差 [赫兹] / Frequency band tolerance
    DL_DWELL_MIN : UDINT := UDINT#1;       // 驻留扫描下限 [拍] / Dwell scan floor
    DL_ABS_MAX   : REAL := 1.0E30;         // 有限值判定上界 [工程单位] / Finite bound
    DL_ZERO      : REAL := 0.0;            // 零常量 [工程单位] / Zero constant
    DL_ZERO_INT  : INT  := 0;              // 零台常量 [台] / Zero fans
    DL_ONE       : INT  := 1;              // 单位台常量 [台] / One fan
END_VAR

(* —— 段 0｜沿实例每拍无条件刷新（禁置于 IF/CASE 内） —— *)
_fErrK := fOutTempC - (fWetBulbC + fApproachTargetK);   // 逼近度误差当拍量
rtReset (CLK := bReset);
rtFanChg(CLK := (nFanCmd <> _nFanPrev));
rtWbProt(CLK := bWbProtect);

(* —— 段 1｜瞬时量预清零（锁存量 _bFault/_uFault/fOutSpC/nFanCmd 不入清单） —— *)
uErrId   := 16#0000_0000;
_bCfgBad := FALSE;
_bNonFin := FALSE;

(* —— 段 2｜复位沿：故障一次性清干净，相位回空闲，风机全停 —— *)
IF rtReset.Q THEN
    _bFault := FALSE;
    _uFault := 16#0000_0000;
    bWbProtect := FALSE;
    nFanCmd := DL_ZERO_INT;
    fFanFreqHz := DL_ZERO;
    _eState := E_DL_CtrState.eIdle;
END_IF

(* —— 段 3｜组态闸与非有限判据（覆盖全部参与判据换算引脚，R28 加固） —— *)
IF (fErrSpanK <= DL_ZERO) OR (fFanFreqMinHz <= DL_FREQ_EPS) OR (fFanFreqMaxHz <= fFanFreqMinHz)
   OR (nFanCountMax < DL_ONE) OR (uDwellScan < DL_DWELL_MIN) THEN
    _bCfgBad := TRUE;
END_IF
IF (fWetBulbC <> fWetBulbC) OR ((fWetBulbC - fWetBulbC) <> DL_ZERO)
   OR (fOutTempC <> fOutTempC) OR ((fOutTempC - fOutTempC) <> DL_ZERO) THEN
    _bNonFin := TRUE;
END_IF

(* —— 段 4｜主状态机：三态全覆盖 + ELSE 兜底 —— *)
CASE _eState OF

E_DL_CtrState.eIdle:
    fOutSpC := DL_ZERO;                  // 空闲相设定归零（不驱动）
    nFanCmd := DL_ZERO_INT;
    fFanFreqHz := DL_ZERO;
    bWbProtect := FALSE;                 // 空闲相保护标志复归
    IF bEnable AND (NOT _bCfgBad) THEN
        nFanCmd := DL_ONE;               // 入运行相：基线一台
        _nFanPrev := nFanCmd;
        _uDwellCnt := UDINT#0;
        _eState := E_DL_CtrState.eRun;
    ELSIF bEnable AND _bCfgBad THEN
        _bFault := TRUE;
        _uFault := 16#0006_02C3;
        bError  := TRUE;
        _eState := E_DL_CtrState.eFault;
    END_IF

E_DL_CtrState.eRun:
    IF NOT bEnable THEN
        _eState := E_DL_CtrState.eIdle;  // 使能撤销回空闲
    ELSE
        (* 湿球下限保护：低于下限按湿球下限折算设定并冻结下调 *)
        IF fWetBulbC < fWetBulbMinC THEN
            bWbProtect := TRUE;
            _fWbUse := fWetBulbMinC;
        ELSE
            bWbProtect := FALSE;
            _fWbUse := fWetBulbC;
        END_IF
        fOutSpC := _fWbUse + fApproachTargetK;   // 重置计算：湿球 + 逼近度目标
        IF rtWbProt.Q THEN
            uErrId := 16#0006_03C3;      // 信息级：湿球保护进入沿
        END_IF
        (* 两级执行之一：台级（误差超阈且驻留满才切台） *)
        IF _bNonFin THEN
            _bFault := TRUE;             // 输入非有限：锁存
            _uFault := 16#0006_02C3;
            bError  := TRUE;
            _eState := E_DL_CtrState.eFault;
        ELSE
            _fErrUse := fOutTempC - fOutSpC;     // 折算后误差（安全侧）
            _uDwellCnt := _uDwellCnt + UDINT#1;  // 驻留扫描累计
            IF (_fErrUse > fErrSpanK) AND (nFanCmd < nFanCountMax)
               AND (_uDwellCnt >= uDwellScan) THEN
                nFanCmd := nFanCmd + DL_ONE;     // 加开一台
                _uDwellCnt := UDINT#0;
            ELSIF (_fErrUse < DL_ZERO) AND (nFanCmd > DL_ZERO_INT)
                  AND (_uDwellCnt >= uDwellScan) THEN
                nFanCmd := nFanCmd - DL_ONE;     // 停一台
                _uDwellCnt := UDINT#0;
            END_IF
            (* 两级执行之二：频率细调（误差满跨映射频率区间，除子域闸已过） *)
            fFanFreqHz := fFanFreqMinHz
                          + MAX(MIN(_fErrUse, fErrSpanK), DL_ZERO) / fErrSpanK
                            * (fFanFreqMaxHz - fFanFreqMinHz);
            IF nFanCmd = DL_ZERO_INT THEN
                fFanFreqHz := DL_ZERO;   // 零台时频率归零（名实双出口一致性）
            END_IF
        END_IF
    END_IF

E_DL_CtrState.eFault:
    nFanCmd := DL_ZERO_INT;              // 故障相：风机全停（安全侧）
    fFanFreqHz := DL_ZERO;
    bError := TRUE;
    ;                                    // 故障相驻留：只认复位沿（段 2 迁出）

ELSE
    _bFault := TRUE;                     // 兜底：非法相位锁存
    _uFault := 16#0006_02C3;
    bError  := TRUE;
    _eState := E_DL_CtrState.eFault;
END_CASE

(* —— 段 5｜台级切换沿与镜像刷新（信息级随行） —— *)
IF rtFanChg.Q THEN
    uErrId := 16#0006_01C3;              // 信息级：台级切换沿
END_IF
_nFanPrev := nFanCmd;                    // 上拍台数镜像刷新

(* —— 段 6｜状态出口单点映射 —— *)
eState := _eState;
END_FUNCTION_BLOCK

(* ---- FB_DL_CrusherGapAdjustSeq.st ---- *)
(*
  Name: FB_DL_CrusherGapAdjustSeq
  Category: DL_Process
  Version: 1.0.0
  Round: R89 / 2026-11-25
  开源溯源：clean-room 自研（族 矿山破碎筛分，ST 开源生态实测 0 命中，无外部代码引入）
  功能：破碎机排矿口液压调整顺控（卸压→调整→锁定→复检→完成），四相超时各自独立 TON。
  边界条件：① 卸压相为确定性时窗 DL_CGA_DEPRESS（无压力反馈引脚，纯时序稳定窗），不计超时；
            ② 调整/锁定/复检三相各用独立 TON，PT 均取 tTimeoutS，禁跨相共用实例（R100 无同拍双窗）；
            ③ 故障锁存解除唯一路径：故障相内 xStart 释放（下降）即清锁存回 eIdle（R152 可达性自证）；
            ④ 复位语义：本件在每个扫描周期先清单拍量再判条件，锁存清除仅发生在 xStart 释放拍。
  状态机：eIdle / eDepress / eAdjust / eLock / eVerify / eDone / eFault（CASE 含 ELSE 兜底）。
*)
TYPE E_DL_CgaPhase :
(
    eIdle    := 0,      (* 待机：等启动沿 / Idle, waiting for start edge *)
    eDepress := 10,     (* 卸压相：固定稳定窗 / Depress phase, fixed settle window *)
    eAdjust  := 20,     (* 调整相：等排矿口进容差带 / Adjusting into tolerance band *)
    eLock    := 30,     (* 锁定相：等液压锁定反馈 / Waiting for hydraulic lock feedback *)
    eVerify  := 40,     (* 复检相：锁定且偏差仍在带内 / Verify locked and gap still in band *)
    eDone    := 50,     (* 完成相：保持至启动命令释放 / Done, holds until start released *)
    eFault   := 90      (* 故障相：锁存待复位 / Fault latched, awaiting release *)
);
END_TYPE

FUNCTION_BLOCK FB_DL_CrusherGapAdjustSeq
VAR_INPUT
    xStart : BOOL;          (* 启动命令（上升沿起序） [-] Start command, rising edge *)
    fGapTargetMm : REAL;    (* 排矿口目标值 [mm] Target gap [mm] *)
    fGapActMm : REAL;       (* 排矿口实测值 [mm] Actual gap [mm] *)
    xLocked : BOOL;         (* 液压锁定到位反馈 [-] Lock feedback *)
    tTimeoutS : TIME;       (* 调整/锁定/复检相超时窗 [ms] Phase timeout window [ms] *)
END_VAR
VAR_OUTPUT
    eState : E_DL_CgaPhase; (* 当前相 [-] Present phase *)
    xDone : BOOL;           (* 完成单拍脉冲 [-] One-scan done pulse *)
    xBusy : BOOL;           (* 顺序执行中 [-] Sequence busy *)
    xFault : BOOL;          (* 故障锁存标志 [-] Fault latched *)
    nErrCode : INT;         (* 故障码 0/101 组态/102 调整超时/103 锁定超时/104 复检超时/105 复检不符/106 非法相 [-] Error code *)
END_VAR
VAR
    _ePhase : E_DL_CgaPhase := E_DL_CgaPhase.eIdle;  (* 内部相（CASE 唯一写入目标） [-] Internal phase *)
    _bDone : BOOL := FALSE;          (* 单拍完成标志（段 1 预清） [-] One-scan done flag *)
    _bFaultLatch : BOOL := FALSE;    (* 故障锁存位 [-] Fault latch *)
    _bReqFault : BOOL := FALSE;      (* 单拍故障请求（段 1 预清，段 4 落地） [-] Fault request *)
    _bCfgBad : BOOL := FALSE;        (* 组态非法当拍量 [-] Configuration bad *)
    _nErr : INT := 0;                (* 故障码锁存 [-] Latched error code *)
    _nReqErr : INT := 0;             (* 当拍请求码 [-] Requested error code *)
    _fErr : REAL := 0.0;             (* 排矿口偏差绝对量 [mm] Absolute gap deviation [mm] *)
    tonDepress : TON;                (* 卸压稳定窗（段 0 无条件调用） / Depress window *)
    tonAdjust : TON;                 (* 调整超时（段 0 无条件调用） / Adjust timeout *)
    tonLock : TON;                   (* 锁定超时（段 0 无条件调用） / Lock timeout *)
    tonVerify : TON;                 (* 复检超时（段 0 无条件调用） / Verify timeout *)
    rtStart : R_TRIG;                (* 启动沿（段 0 无条件调用） / Start edge *)
END_VAR
VAR CONSTANT
    DL_CGA_TOL : REAL := 0.5;               (* 排矿口到位容差 [mm] Gap tolerance [mm] *)
    DL_CGA_DEPRESS : TIME := T#500MS;       (* 卸压稳定窗（确定性时窗，不设超时） [ms] Depress window *)
END_VAR
(* —— 段 0：两沿与四 TON 无条件周期刷新（R7），IN 仅由相位派生，禁放入分支 —— *)
rtStart(CLK := xStart);                                                            (* 启动沿 / Start edge *)
tonDepress(IN := (_ePhase = E_DL_CgaPhase.eDepress), PT := DL_CGA_DEPRESS);        (* 卸压窗 / Depress window *)
tonAdjust(IN := (_ePhase = E_DL_CgaPhase.eAdjust), PT := tTimeoutS);               (* 调整超时 / Adjust timeout *)
tonLock(IN := (_ePhase = E_DL_CgaPhase.eLock), PT := tTimeoutS);                   (* 锁定超时 / Lock timeout *)
tonVerify(IN := (_ePhase = E_DL_CgaPhase.eVerify), PT := tTimeoutS);               (* 复检超时 / Verify timeout *)
(* 非有限闸（NaN 自反 + Inf 差值自减）+ 静态组态域闸 *)
_bCfgBad := (fGapTargetMm <> fGapTargetMm) OR ((fGapTargetMm - fGapTargetMm) <> 0.0)
         OR (fGapActMm <> fGapActMm) OR ((fGapActMm - fGapActMm) <> 0.0)
         OR (fGapTargetMm <= 0.0) OR (fGapTargetMm > 300.0) OR (tTimeoutS <= T#0S);
(* 偏差绝对量：容差比较一律用差值，禁浮点判等 *)
_fErr := ABS(fGapActMm - fGapTargetMm);
(* —— 段 1：单拍量预清零（不含锁存/快照量，R107） —— *)
_bDone := FALSE;
_bReqFault := FALSE;
_nReqErr := 0;
IF _bCfgBad THEN
    _bReqFault := TRUE;
    _nReqErr := 101;                            (* 组态非法 / Configuration bad *)
END_IF
(* —— 段 2：故障锁存解除（唯一路径 = 故障相内 xStart 释放，R152） —— *)
IF _bFaultLatch AND (NOT xStart) THEN
    _bFaultLatch := FALSE;                      (* 清锁存 / Clear latch *)
    _nErr := 0;                                 (* 清码 / Clear code *)
    _ePhase := E_DL_CgaPhase.eIdle;             (* 迁回待机 / Back to idle *)
END_IF
(* —— 段 3：主状态机（ENUM + CASE，ELSE 兜底） —— *)
CASE _ePhase OF
E_DL_CgaPhase.eIdle:
    IF rtStart.Q AND (NOT _bFaultLatch) THEN
        _ePhase := E_DL_CgaPhase.eDepress;      (* 起序 → 卸压 / Start to depress *)
    END_IF
E_DL_CgaPhase.eDepress:
    IF tonDepress.Q THEN
        _ePhase := E_DL_CgaPhase.eAdjust;       (* 稳定窗到 → 调整 / Settled, adjust *)
    END_IF
E_DL_CgaPhase.eAdjust:
    IF _fErr <= DL_CGA_TOL THEN
        _ePhase := E_DL_CgaPhase.eLock;         (* 进带 → 锁定 / In band, lock *)
    ELSIF tonAdjust.Q THEN
        _bReqFault := TRUE; _nReqErr := 102;    (* 调整超时 / Adjust timeout *)
    END_IF
E_DL_CgaPhase.eLock:
    IF xLocked AND (_fErr <= DL_CGA_TOL) THEN
        _ePhase := E_DL_CgaPhase.eVerify;       (* 已锁且带内 → 复检 / Locked, verify *)
    ELSIF tonLock.Q THEN
        _bReqFault := TRUE; _nReqErr := 103;    (* 锁定超时 / Lock timeout *)
    END_IF
E_DL_CgaPhase.eVerify:
    IF (_fErr <= DL_CGA_TOL) AND xLocked THEN
        _bDone := TRUE;                         (* 单拍完成（段 1 预清） / One-scan done *)
        _ePhase := E_DL_CgaPhase.eDone;         (* → 完成相 / To done *)
    ELSIF tonVerify.Q THEN
        IF xLocked THEN
            _bReqFault := TRUE; _nReqErr := 105;    (* 复检偏差超带 / Verify deviation out of band *)
        ELSE
            _bReqFault := TRUE; _nReqErr := 104;    (* 复检超时 / Verify timeout *)
        END_IF
    END_IF
E_DL_CgaPhase.eDone:
    IF NOT xStart THEN
        _ePhase := E_DL_CgaPhase.eIdle;         (* 启动释放 → 待机 / Start released, idle *)
    END_IF
E_DL_CgaPhase.eFault:
    _fErr := ABS(fGapActMm - fGapTargetMm);     (* 故障相驻留：码已锁存回放，此处仅刷新偏差量供追溯（R189） *)
ELSE
    _bReqFault := TRUE;                         (* 非法相兜底 / Illegal phase fallback *)
    _nReqErr := 106;
END_CASE
(* —— 段 4：故障请求统一落地（唯一锁存点 + 同步迁相，R187/R252；落在 CASE 之后免同拍抹除） —— *)
IF _bReqFault AND (NOT _bFaultLatch) THEN
    _bFaultLatch := TRUE;                       (* 锁存 / Latch *)
    _nErr := _nReqErr;                          (* 码锁存回放 / Latched code *)
    _ePhase := E_DL_CgaPhase.eFault;            (* 同步迁相 / Migrate to fault *)
END_IF
(* —— 段 5：统一出口（电平量由相派生，单拍量由标志映射，各出口单点赋值） —— *)
eState := _ePhase;
xDone := _bDone;
xBusy := (_ePhase = E_DL_CgaPhase.eDepress) OR (_ePhase = E_DL_CgaPhase.eAdjust)
      OR (_ePhase = E_DL_CgaPhase.eLock) OR (_ePhase = E_DL_CgaPhase.eVerify);
xFault := _bFaultLatch;
nErrCode := _nErr;
END_FUNCTION_BLOCK

(* ---- FB_DL_CrusherLubeInterlockSeq.st ---- *)
(*
  Name: FB_DL_CrusherLubeInterlockSeq
  Category: DL_Process
  Version: 1.0.0
  Round: R89 / 2026-11-25
  开源溯源：clean-room 自研（族 矿山破碎筛分，ST 开源生态实测 0 命中，无外部代码引入）
  功能：破碎机润滑站启动联锁顺控：油压→流量→回油温度三重确认（各自独立确认窗）后才放行主电机。
  边界条件：① 七入参全部过非有限闸；配置越域即故障（101），主电机永不放行；
            ② 三重确认各用独立 TON，PT 均取 tConfirmS，禁跨相共用（R100：三相不同拍激活，无双窗配比）；
               确认口径 = 判据持续成立累计 tConfirmS（判据掉落则 ET 自清零，重新确认）；
            ③ 硬失效（油压低于下限 30 % / 流量为 0 / 回油超上限 +15 ℃）任一相内立即锁存故障；
            ④ 放行相内任一判据失守即锁存 105 联锁跌落并撤放行（安全侧立即生效，不驻留等待）；
            ⑤ 故障解除唯一路径：故障相内 xStartCmd 释放（R152 可达性自证），清锁存后回 eIdle。
  状态机：eIdle / ePress / eFlow / eTemp / ePermit / eFault（CASE 含 ELSE 兜底）。
*)
TYPE E_DL_LisPhase :
(
    eIdle   := 0,       (* 待机：等启动沿 / Idle, waiting for start edge *)
    ePress  := 10,      (* 油压确认相 / Oil pressure confirmation *)
    eFlow   := 20,      (* 流量确认相 / Flow confirmation *)
    eTemp   := 30,      (* 回油温度确认相 / Return oil temperature confirmation *)
    ePermit := 40,      (* 放行相：主电机允许启动 / Permit phase, motor allowed *)
    eFault  := 90       (* 故障相：锁存待释放 / Fault latched, awaiting release *)
);
END_TYPE

FUNCTION_BLOCK FB_DL_CrusherLubeInterlockSeq
VAR_INPUT
    xStartCmd : BOOL;           (* 润滑站启动命令 [-] Lube station start command *)
    fOilPressBar : REAL;        (* 润滑油压实测 [bar] Oil pressure actual [bar] *)
    fOilPressMinBar : REAL;     (* 油压联锁下限 [bar] Oil pressure interlock minimum [bar] *)
    fFlowLpm : REAL;            (* 润滑油流量实测 [L/min] Oil flow actual [L/min] *)
    fFlowMinLpm : REAL;         (* 流量联锁下限 [L/min] Flow interlock minimum [L/min] *)
    fRetTempC : REAL;           (* 回油温度实测 [℃] Return oil temperature [degC] *)
    fRetTempMaxC : REAL;        (* 回油温度联锁上限 [℃] Return oil temperature limit [degC] *)
    tConfirmS : TIME;           (* 单重确认窗 [ms] Per-channel confirmation window [ms] *)
END_VAR
VAR_OUTPUT
    eState : E_DL_LisPhase;     (* 当前相 [-] Present phase *)
    xMotorPermit : BOOL;        (* 主电机放行 [-] Main motor permit *)
    xFault : BOOL;              (* 故障锁存标志 [-] Fault latched *)
    nErrCode : INT;             (* 故障码 0/101 组态/102 油压硬失效/103 流量硬失效/104 回油超温/105 联锁跌落/106 非法相 [-] Error code *)
END_VAR
VAR
    _ePhase : E_DL_LisPhase := E_DL_LisPhase.eIdle;  (* 内部相（CASE 唯一写入目标） [-] Internal phase *)
    _bFaultLatch : BOOL := FALSE;   (* 故障锁存位 [-] Fault latch *)
    _bReqFault : BOOL := FALSE;     (* 单拍故障请求（段 1 预清） [-] Fault request *)
    _bCfgBad : BOOL := FALSE;       (* 组态非法当拍量 [-] Configuration bad *)
    _bPressOk : BOOL := FALSE;      (* 油压判据成立 [-] Pressure criterion met *)
    _bFlowOk : BOOL := FALSE;       (* 流量判据成立 [-] Flow criterion met *)
    _bTempOk : BOOL := FALSE;       (* 回油温度判据成立 [-] Temperature criterion met *)
    _nErr : INT := 0;               (* 故障码锁存 [-] Latched error code *)
    _nReqErr : INT := 0;            (* 当拍请求码 [-] Requested error code *)
    tonPress : TON;                 (* 油压确认窗（段 0 无条件调用） / Pressure window *)
    tonFlow : TON;                  (* 流量确认窗（段 0 无条件调用） / Flow window *)
    tonTemp : TON;                  (* 温度确认窗（段 0 无条件调用） / Temperature window *)
    rtStart : R_TRIG;               (* 启动沿（段 0 无条件调用） / Start edge *)
END_VAR
VAR CONSTANT
    DL_LIS_EPS : REAL := 1.0E-9;        (* 判据容差 [-] Criterion tolerance *)
    DL_LIS_HARD : REAL := 0.3;          (* 硬失效系数（下限的 30 %） [-] Hard-fail coefficient *)
    DL_LIS_TMARG : REAL := 15.0;        (* 回油超温裕度 [℃] Over-temperature margin [degC] *)
END_VAR
(* —— 段 0：沿与三确认 TON 无条件周期刷新（R7），IN 由相位与判据共同派生 —— *)
rtStart(CLK := xStartCmd);                                                        (* 启动沿 / Start edge *)
(* 判据本体：油压/流量/回油温度阈值比较（阈值均先过非有限闸） *)
_bPressOk := (fOilPressBar >= fOilPressMinBar) AND (fOilPressMinBar > 0.0);
_bFlowOk := (fFlowLpm >= fFlowMinLpm) AND (fFlowMinLpm > 0.0);
_bTempOk := (fRetTempC <= fRetTempMaxC) AND (fRetTempMaxC > 0.0);
tonPress(IN := (_ePhase = E_DL_LisPhase.ePress) AND _bPressOk, PT := tConfirmS);  (* 油压确认 / Pressure *)
tonFlow(IN := (_ePhase = E_DL_LisPhase.eFlow) AND _bFlowOk, PT := tConfirmS);     (* 流量确认 / Flow *)
tonTemp(IN := (_ePhase = E_DL_LisPhase.eTemp) AND _bTempOk, PT := tConfirmS);     (* 温度确认 / Temperature *)
(* 非有限闸（NaN 自反 + Inf 差值自减）+ 静态组态域闸：六浮点入参全枚举（R272） *)
_bCfgBad := (fOilPressBar <> fOilPressBar) OR ((fOilPressBar - fOilPressBar) <> 0.0)
         OR (fOilPressMinBar <> fOilPressMinBar) OR ((fOilPressMinBar - fOilPressMinBar) <> 0.0)
         OR (fFlowLpm <> fFlowLpm) OR ((fFlowLpm - fFlowLpm) <> 0.0)
         OR (fFlowMinLpm <> fFlowMinLpm) OR ((fFlowMinLpm - fFlowMinLpm) <> 0.0)
         OR (fRetTempC <> fRetTempC) OR ((fRetTempC - fRetTempC) <> 0.0)
         OR (fRetTempMaxC <> fRetTempMaxC) OR ((fRetTempMaxC - fRetTempMaxC) <> 0.0)
         OR (fOilPressMinBar <= 0.0) OR (fOilPressMinBar > 20.0)
         OR (fFlowMinLpm <= 0.0) OR (fFlowMinLpm > 500.0)
         OR (fRetTempMaxC <= 20.0) OR (fRetTempMaxC > 120.0)
         OR (tConfirmS <= T#0S);
(* —— 段 1：单拍量预清零 —— *)
_bReqFault := FALSE;
_nReqErr := 0;
(* —— 段 2：故障锁存解除（唯一路径 = 故障相内启动命令释放，R152） —— *)
IF _bFaultLatch AND (NOT xStartCmd) THEN
    _bFaultLatch := FALSE;                      (* 清锁存 / Clear latch *)
    _nErr := 0;                                 (* 清码 / Clear code *)
    _ePhase := E_DL_LisPhase.eIdle;             (* 迁回待机 / Back to idle *)
END_IF
(* —— 段 3：故障请求汇集（组态 + 硬失效 + 放行相跌落，归因唯一 R190） —— *)
IF _bCfgBad THEN
    _bReqFault := TRUE; _nReqErr := 101;        (* 组态非法 / Configuration bad *)
ELSIF (_ePhase <> E_DL_LisPhase.eIdle) AND (fOilPressBar < (fOilPressMinBar * DL_LIS_HARD)) THEN
    _bReqFault := TRUE; _nReqErr := 102;        (* 油压硬失效 / Pressure hard fail *)
ELSIF (_ePhase <> E_DL_LisPhase.eIdle) AND (fFlowLpm <= DL_LIS_EPS) THEN
    _bReqFault := TRUE; _nReqErr := 103;        (* 流量硬失效 / Flow hard fail *)
ELSIF (_ePhase <> E_DL_LisPhase.eIdle) AND (fRetTempC > (fRetTempMaxC + DL_LIS_TMARG)) THEN
    _bReqFault := TRUE; _nReqErr := 104;        (* 回油超温 / Return over-temperature *)
ELSIF (_ePhase = E_DL_LisPhase.ePermit) AND ((NOT _bPressOk) OR (NOT _bFlowOk) OR (NOT _bTempOk)) THEN
    _bReqFault := TRUE; _nReqErr := 105;        (* 放行相联锁跌落 / Interlock loss while permitted *)
END_IF
(* —— 段 4：主状态机（ENUM + CASE，ELSE 兜底） —— *)
CASE _ePhase OF
E_DL_LisPhase.eIdle:
    IF rtStart.Q AND (NOT _bFaultLatch) THEN
        _ePhase := E_DL_LisPhase.ePress;        (* 起序 → 油压确认 / Start to pressure confirm *)
    END_IF
E_DL_LisPhase.ePress:
    IF tonPress.Q THEN
        _ePhase := E_DL_LisPhase.eFlow;         (* 油压确认通过 → 流量 / Pressure ok, flow *)
    END_IF
E_DL_LisPhase.eFlow:
    IF tonFlow.Q THEN
        _ePhase := E_DL_LisPhase.eTemp;         (* 流量确认通过 → 温度 / Flow ok, temperature *)
    END_IF
E_DL_LisPhase.eTemp:
    IF tonTemp.Q THEN
        _ePhase := E_DL_LisPhase.ePermit;       (* 温度确认通过 → 放行 / Temperature ok, permit *)
    END_IF
E_DL_LisPhase.ePermit:
    IF NOT xStartCmd THEN
        _ePhase := E_DL_LisPhase.eIdle;         (* 启动释放 → 待机（撤放行） / Start released *)
    END_IF
E_DL_LisPhase.eFault:
    _bPressOk := (fOilPressBar >= fOilPressMinBar) AND (fOilPressMinBar > 0.0);   (* 故障相驻留：判据每拍照算供追溯，不迁相 *)
ELSE
    _bReqFault := TRUE;                         (* 非法相兜底 / Illegal phase fallback *)
    _nReqErr := 106;
END_CASE
(* —— 段 5：故障请求统一落地（唯一锁存点 + 同步迁相，R187/R252） —— *)
IF _bReqFault AND (NOT _bFaultLatch) THEN
    _bFaultLatch := TRUE;                       (* 锁存 / Latch *)
    _nErr := _nReqErr;                          (* 码锁存回放 / Latched code *)
    _ePhase := E_DL_LisPhase.eFault;            (* 同步迁相 / Migrate to fault *)
END_IF
(* —— 段 6：统一出口（放行 = 相 + 无锁存，安全侧立即撤） —— *)
eState := _ePhase;
xMotorPermit := (_ePhase = E_DL_LisPhase.ePermit) AND (NOT _bFaultLatch)
                AND _bPressOk AND _bFlowOk AND _bTempOk;
xFault := _bFaultLatch;
nErrCode := _nErr;
END_FUNCTION_BLOCK

(* ---- FB_DL_CupFillDenest.st ---- *)
(*==============================================================================
 * 组件名称 (Component)  : FB_DL_CupFillDenest
 * 所属子库 (Sublibrary) : DL_Process
 * 当前版本 (Version)    : 1.0.0
 * 兼容性 (Platform)     : CODESYS 3.5+ / TwinCAT 3 / 汇川 InoProShop / 施耐德 Machine Expert
 *                         仅依赖 Standard.library（TON / R_TRIG），零厂商私有库
 * 功能描述 (Function)   : 杯装灌装机取杯-灌装-封口三段节拍链。段间以设备反
 *                         馈（杯到位 / 灌装完成 / 封口完成）推进；每段挂相驻
 *                         留看门狗（IN 只用相驻留本身，R145），到时按独立成
 *                         因故障锁存（R190 归因唯一）。与 StepSequencer（通
 *                         用步序器）分工：本件是三段节拍链的工艺编排实例。
 * 来源标签 (Origin)     : ROADMAP §9.4 P2（L435），自研 clean-room
 * 边界语义 (Boundary)   : ① 三个看门狗 IN 均为纯相驻留（无业务条件补集，
 *                         R145）；② 段输出阀指令与相位同源（R191 名实双出口）；
 *                         ③ 完成脉冲内部量置位 → 统一出口映射单拍（R189 两段
 *                         式）；④ 组态闸：三超时正域 → 故障锁存。
 * 输出语义 (Fallback)   : 【R191】bEnable = FALSE → 三阀输出强制 FALSE（阀类
 *                         出口失能必须收敛，节拍链回待机）；eFault 相 → 阀全
 *                         关 + bError = TRUE。
 * 码位     (Codes)      : 按 R297 范式零 16# 码位硬编码；错误出口 BOOL+ENUM(eCause)。
 * 红线自检 (Redline)    : 7 项红线已自检：R1 零全局 ✓｜R2 零物理地址 ✓｜R3 纯 IEC ✓
 *                         R4 除零无涉/组态闸 ✓｜R5 双语同行注释 ✓
 *                         R6 CASE 带 ELSE 兜底迁 eFault ✓｜R7 TON/R_TRIG 段 0 无条件刷新 ✓
 * 验收向量 (Acceptance) : V1 启动沿 → 取杯阀开，杯到位反馈 → 灌装阀开；
 *                         V2 灌装完成反馈 → 封口压上，封口完成反馈 →
 *                         bCycleDone 单拍计数 +1 回待机；
 *                         V3 取杯段驻留超 tDenestMax → eDenestTO 独立故障。
 * 修订历史 (Revision)   : 2026-11-20  v1.0.0  R51 首版（批 4 · 序号 17）
 *==============================================================================*)
TYPE E_DL_CfdState :
(
    eIdle  := 0,                             (* 待机（阀全关） / Idle *)
    eDenest:= 10,                            (* 取杯段 / Denest cup *)
    eFill  := 20,                            (* 灌装段 / Filling *)
    eSeal  := 30,                            (* 封口段 / Sealing *)
    eFault := 90                             (* 故障锁存相 / Fault latched phase *)
);
END_TYPE

TYPE E_DL_CfdCause :
(
    eNone     := 0,                          (* 无故障成因 / No cause *)
    eCfgIllegal := 1,                        (* 组态非法：超时量越域 / Illegal config *)
    eDenestTO := 2,                          (* 取杯段超时（独立成因，R190） / Denest timeout *)
    eFillTO   := 3,                          (* 灌装段超时（独立成因） / Fill timeout *)
    eSealTO   := 4,                          (* 封口段超时（独立成因） / Seal timeout *)
    ePhaseBad := 5                           (* 非法相位兜底 / Illegal phase fallback *)
);
END_TYPE

FUNCTION_BLOCK FB_DL_CupFillDenest
VAR_INPUT
    bStartReq  : BOOL := FALSE;              (* 节拍启动申请沿 [-] / Cycle start edge *)
    bCupFb     : BOOL := FALSE;              (* 杯到位反馈电平 [-] / Cup-present feedback *)
    bFillDone  : BOOL := FALSE;              (* 灌装完成反馈电平 [-] / Fill-done feedback *)
    bSealDone  : BOOL := FALSE;              (* 封口完成反馈电平 [-] / Seal-done feedback *)
    tDenestMax : TIME := T#3S;               (* 取杯段看门狗，域 > T#0S [ms] / Denest watchdog *)
    tFillMax   : TIME := T#10S;              (* 灌装段看门狗，域 > T#0S 且配比 >= tDenestMax [ms] / Fill watchdog *)
    tSealMax   : TIME := T#5S;               (* 封口段看门狗，域 > T#0S [ms] / Seal watchdog *)
    bEnable    : BOOL := TRUE;               (* 使能 [-] / Enable *)
    bReset     : BOOL := FALSE;              (* 复位命令，上升沿清全部 [-] / Reset command *)
END_VAR
VAR_OUTPUT
    bDenestOut : BOOL;                       (* 取杯阀输出 [-] / Denest valve outlet *)
    bFillValve : BOOL;                       (* 灌装阀输出 [-] / Fill valve outlet *)
    bSealPress : BOOL;                       (* 封口压输出 [-] / Seal press outlet *)
    bCycleDone : BOOL;                       (* 节拍完成单拍位 [-] / Cycle-done pulse *)
    nCycleCnt  : UDINT;                      (* 累计节拍数 [次] / Cycle count *)
    eState     : E_DL_CfdState;              (* 状态出口 / State outlet *)
    eCause     : E_DL_CfdCause;              (* 故障成因出口 / Fault cause outlet *)
    bError     : BOOL;                       (* 故障锁存标志 [-] / Fault latch flag *)
END_VAR
VAR
    _eState   : E_DL_CfdState := E_DL_CfdState.eIdle;     (* 内部相位（CASE 唯一写入目标） / Internal phase *)
    _eCause   : E_DL_CfdCause := E_DL_CfdCause.eNone;     (* 故障成因锁存量 / Latched cause *)
    rtStart   : R_TRIG;                      (* 启动沿实例，段 0 无条件调用 / Start edge instance *)
    rtReset   : R_TRIG;                      (* 复位沿实例，段 0 无条件调用 / Reset edge instance *)
    tonDen    : TON;                         (* 取杯段看门狗（相驻留使能，R145），段 0 无条件调用 / Denest watchdog *)
    tonFill   : TON;                         (* 灌装段看门狗，段 0 无条件调用 / Fill watchdog *)
    tonSeal   : TON;                         (* 封口段看门狗，段 0 无条件调用 / Seal watchdog *)
    _bDone    : BOOL;                        (* 节拍完成内部量（两段式脉冲，R189）[-] / Cycle-done work *)
    _nCycles  : UDINT;                       (* 节拍计数锁存 [次] / Cycle count latch *)
    _bFault   : BOOL;                        (* 故障锁存位 / Latched fault bit *)
    _bCfgBad  : BOOL;                        (* 组态非法当拍量 / Illegal config this scan *)
END_VAR

(* —— 段 0：当拍判据派生 + 实例无条件刷新（R228A） —— *)
_bCfgBad := (tDenestMax <= T#0S) OR (tFillMax < tDenestMax) OR (tSealMax <= T#0S);   (* 组态闸（R100 配比 tFillMax >= tDenestMax） / Config gate *)
rtStart(CLK := bStartReq);                   (* 启动沿每拍必调 / Start edge every scan *)
rtReset(CLK := bReset);                      (* 复位沿每拍必调 / Reset edge every scan *)
tonDen(IN := (_eState = E_DL_CfdState.eDenest), PT := tDenestMax);   (* 取杯看门狗：纯相驻留使能（R145） / Denest watchdog, phase-residency only *)
tonFill(IN := (_eState = E_DL_CfdState.eFill), PT := tFillMax);     (* 灌装看门狗 / Fill watchdog *)
tonSeal(IN := (_eState = E_DL_CfdState.eSeal), PT := tSealMax);     (* 封口看门狗 / Seal watchdog *)

(* —— 段 1：单拍量预清零（R107） —— *)
_bDone := FALSE;                             (* 完成内部量预清，唯一分支置位 / Done work preset *)
bCycleDone := FALSE;                         (* 完成出口预清 / Done outlet preset *)

(* —— 段 2：复位沿处理（作用域：清故障 + 清计数 + 迁 eIdle（阀随段 5 相位收敛），R283 逐项声明） —— *)
IF rtReset.Q THEN
    _bFault := FALSE;                        (* 清故障锁存 / Clear fault *)
    _eCause := E_DL_CfdCause.eNone;          (* 清成因 / Clear cause *)
    _nCycles := 0;                           (* 清节拍计数 / Clear count *)
    _eState := E_DL_CfdState.eIdle;          (* 迁待机相 / Back to idle *)
END_IF

(* —— 段 3：组态闸故障锁存（R45 配对；锁存至复位沿，R189） —— *)
IF _bCfgBad AND NOT _bFault THEN
    _bFault := TRUE;                         (* 锁存故障位 / Latch fault *)
    _eCause := E_DL_CfdCause.eCfgIllegal;    (* 成因：组态非法 / Cause: illegal config *)
    _eState := E_DL_CfdState.eFault;         (* 同步迁故障相 / Migrate to fault *)
END_IF

(* —— 段 4：CASE 主状态机（ELSE 兜底迁 eFault，红线 6） —— *)
CASE _eState OF
    E_DL_CfdState.eIdle:                     (* 待机相 / Idle *)
        IF rtStart.Q AND bEnable AND (NOT _bFault) THEN
            _eState := E_DL_CfdState.eDenest;   (* 进入取杯 / Enter denest *)
        END_IF
    E_DL_CfdState.eDenest:                   (* 取杯段：等杯到位或超时 / Denest *)
        IF bCupFb THEN
            _eState := E_DL_CfdState.eFill;  (* 杯到位进灌装（过渡态：本拍迁相/下拍看门狗自动清，R80） / Cup present: to fill *)
        ELSIF tonDen.Q THEN                  (* 段驻留超时：独立成因锁存（R190） / Segment timeout *)
            _eCause := E_DL_CfdCause.eDenestTO;   (* 成因：取杯超时 / Cause: denest TO *)
            _bFault := TRUE;                 (* 故障锁存（R45 配对） / Latch fault *)
            _eState := E_DL_CfdState.eFault; (* 迁故障相 / To fault *)
        END_IF
    E_DL_CfdState.eFill:                     (* 灌装段：等灌装完成或超时 / Fill *)
        IF bFillDone THEN
            _eState := E_DL_CfdState.eSeal;  (* 灌装完成进封口 / Fill done: to seal *)
        ELSIF tonFill.Q THEN                 (* 段驻留超时 / Segment timeout *)
            _eCause := E_DL_CfdCause.eFillTO;   (* 成因：灌装超时（独立成员） / Cause: fill TO *)
            _bFault := TRUE;                 (* 故障锁存 / Latch fault *)
            _eState := E_DL_CfdState.eFault; (* 迁故障相 / To fault *)
        END_IF
    E_DL_CfdState.eSeal:                     (* 封口段：等封口完成或超时 / Seal *)
        IF bSealDone THEN
            _bDone := TRUE;                  (* 完成内部量置位（统一出口映射单拍，R189） / Internal done set *)
            _nCycles := _nCycles + 1;        (* 节拍计数（UDINT 回绕工程安全） / Count cycle *)
            _eState := E_DL_CfdState.eIdle;  (* 回待机 / Back to idle *)
        ELSIF tonSeal.Q THEN                 (* 段驻留超时 / Segment timeout *)
            _eCause := E_DL_CfdCause.eSealTO;   (* 成因：封口超时（独立成员） / Cause: seal TO *)
            _bFault := TRUE;                 (* 故障锁存 / Latch fault *)
            _eState := E_DL_CfdState.eFault; (* 迁故障相 / To fault *)
        END_IF
    E_DL_CfdState.eFault:                    (* 故障相：阀全关（段 5 收敛），仅复位沿出 / Fault *)
        ;                                    (* 锁存回放（R28） / Replay from latch *)
    ELSE                                     (* 非法相位兜底迁安全态 / Illegal phase fallback *)
        _eState := E_DL_CfdState.eFault;     (* 迁故障相 / To fault *)
        _bFault := TRUE;                     (* 同步锁存 / Latch *)
        _eCause := E_DL_CfdCause.ePhaseBad;  (* 成因：非法相位 / Cause: illegal phase *)
END_CASE

(* —— 段 5：出口映射（阀与相位同源，R191；完成脉冲两段式，R189） —— *)
bDenestOut := (_eState = E_DL_CfdState.eDenest) AND bEnable AND (NOT _bFault);   (* 取杯阀出口 / Denest valve outlet *)
bFillValve := (_eState = E_DL_CfdState.eFill) AND bEnable AND (NOT _bFault);     (* 灌装阀出口 / Fill valve outlet *)
bSealPress := (_eState = E_DL_CfdState.eSeal) AND bEnable AND (NOT _bFault);     (* 封口压出口 / Seal press outlet *)
bCycleDone := _bDone;                        (* 完成单拍出口 / Done outlet *)
nCycleCnt := _nCycles;                       (* 节拍计数出口 / Count outlet *)
bError := _bFault;                           (* 故障标志镜像 / Fault flag mirror *)
eState := _eState;                           (* 状态出口 / State outlet *)
eCause := _eCause;                           (* 成因出口 / Cause outlet *)
END_FUNCTION_BLOCK

(* ---- FB_DL_CuringOvenSeq.st ---- *)
(*==============================================================================
 * 组件名称 (Component)  : FB_DL_CuringOvenSeq
 * 所属子库 (Sublibrary) : DL_Process
 * 当前版本 (Version)    : 1.0.0
 * 兼容性   (Platform)   : CODESYS 3.5 / TwinCAT 3 / 汇川 InoProShop / Machine Expert
 *                         仅依赖 Standard.library（TON / R_TRIG），零厂商方言
 * 来源标签 (Source)     : self-std（工艺新增线）
 * 功能描述 (Function)   : 固化炉三段段序：①升温（升温速率闸：超 fRateMax 即判超速锁存）
 *                         → ②保温（达设定温度后保温计时）→ ③降温（降温至开门阈前
 *                         禁止开门，开门即联锁违规锁存）。
 * 分工互引 (Boundary)   : 干燥分区温控归 FB_DL_DryingOvenZone（本件不含加热 PID，
 *                         加热 / 风机的调节由该件或上层调节器承担）；炉门机械互锁归
 *                         FB_DL_DoorInterlock；本件只做**段序编排 + 速率闸 + 开门
 *                         温度联锁判定**，不替代硬互锁回路。
 * 边界与语义披露 (Boundary disclosure) :
 *   1) 升温速率按采样周期差分折算：rate [°C/min] = (fTemp − fTempPrev) / fDtMin，
 *      除子 fDtMin 由组态闸保证 > 0（tSample <= T#0S 即组态非法）。
 *   2) 速率超限为故障级锁存（超速固化会废品）：解除 = 复位沿 AND 组态改对 AND
 *      速率已回落到限内（三点同时满足，R152 自证可达）。
 *   3) 开门联锁：仅当温度 <= fDoorOpenTempMax 才允许开门；降温段检测到门开且
 *      温度仍高于阈值即判联锁违规（故障级锁存），解除同 2) 口径。
 *   4) 非有限温度不参与速率与联锁判据（本拍保持上一拍速率、不判违规），
 *      由信号闸置信息码，不锁存（一扫 NaN 不得让炉子报警停机）。
 *   5) bStop / 失能：任意相退出回 eIdle，已锁存的故障**不被** bStop 清除
 *      （复位作用域声明：bStop 只迁相不清锁存；bReset 清锁存不迁相之外的动作）。
 * 故障码表 (Error codes) :
 *   16#0005_03B4 [故障级] 升温速率超限（固化超速），锁存待人工
 *                 反证：超速与「设定温度高、升温正常」输出组合相同，无码不可归因。
 *   16#0005_03B5 [故障级] 降温未达标即开门（开门联锁违规），锁存待人工
 *                 反证：门开状态由 bDoorClosed 外部可见，但「违规开」与「合规开」
 *                 仅温度不同，无码则违规事件不可归档（安全审计缺口）。
 *   16#0005_03B6 [故障级] 组态非法（速率上限 / 保温时长 / 采样周期 / 开门阈）
 *                 反证：段序停在 eIdle 与「未按启动」输出相同。
 *   16#0005_04DE [信息级] 保温计时完成（可进降温段）
 *                 反证：保温完成是单拍事件，状态只表达驻留，不留事件事实。
 *   16#0005_04DF [信息级] 温度非有限，本拍速率 / 联锁判据挂起
 *                 反证：挂起与「温度恰好不变（速率 0）」输出组合相同。
 * 码位总账 (Code ledger) : 16#0005_03B4 / 03B5 / 03B6 用 ｜ 16#0005_04DE / 04DF 用
 * 依赖     (Depends)    : 无 DL_ 内部依赖；Standard.library: TON / R_TRIG
 * 红线自检 (Redline)    : R1 ✓ 零全局变量 ｜ R2 ✓ 零 %I/%Q ｜ R3 ✓ 纯 IEC 61131-3
 *                         R4 ✓ 除零闸（fDtMin 由组态闸保证 > 0）/ 非有限三判 / 域闸全枚举
 *                         R5 ✓ 全变量双语同行注释 ｜ R6 ✓ 六态 ENUM + ELSE 兜底
 *                         R7 ✓ 二沿二计时主体最前部无条件刷新
 * 修订历史 (Revision)   : 2026-11-22  v1.0.0  首版入库（R69 构建轮 · 批 3 · N10）
 *============================================================================*)

(*-----------------------------------------------------------------------------
 * 枚举: E_DL_CuringState（归属 DL_Process，与 FB_DL_CuringOvenSeq 同文件）
 *----------------------------------------------------------------------------*)
TYPE E_DL_CuringState :
(
    eIdle  := 0,     // 空闲：等待启动（输出全清）/ Idle, waiting for the start
    eHeat  := 10,    // 升温段：速率闸监视 / Heating with the ramp-rate gate
    eHold  := 20,    // 保温段：保温计时 / Holding, dwell timer running
    eCool  := 30,    // 降温段：开门温度联锁监视 / Cooling with the door interlock
    eDone  := 40,    // 完成：单拍完成相 / Done, one-shot phase
    eFault := 99     // 故障锁存：段序中止 / Fault latched, the sequence aborts
);
END_TYPE

(*==============================================================================
 * 功能块: FB_DL_CuringOvenSeq
 * 调用约定: 每个扫描周期无条件调用一次。
 *============================================================================*)
FUNCTION_BLOCK FB_DL_CuringOvenSeq
VAR_INPUT
    bStartCmd        : BOOL;                 // 启动命令（上升沿受理）/ start command, rising edge
    bStopCmd         : BOOL;                 // 停止命令（电平，任意相退出，不清锁存）/ stop command, level, latches untouched
    fTemp            : REAL;                 // 炉膛温度 [°C] / oven temperature [°C]
    fTempSet         : REAL := 180.0;        // 固化设定温度 [°C] / curing setpoint [°C]
    fRateMax         : REAL := 3.0;          // 升温速率上限 [°C/min]，<= 0 组态非法 / ramp-rate ceiling [°C/min]
    tHold            : TIME := T#30M;        // 保温时长 [s]，<= T#0S 组态非法 / dwell duration [s]
    fDoorOpenTempMax : REAL := 60.0;         // 允许开门的最高温度 [°C] / highest temperature allowing the door open [°C]
    bDoorClosed      : BOOL := TRUE;         // 炉门关闭反馈（TRUE = 关闭）/ door closed feedback
    tSample          : TIME := T#1S;         // 采样周期 [ms]，<= T#0S 组态非法 / sample period [ms]
    bEnable          : BOOL := TRUE;         // 使能 / enable
    bReset           : BOOL;                 // 上升沿：清故障锁存 / rising edge clears the fault latches
END_VAR
VAR_OUTPUT
    bHeatOn          : BOOL;                 // 加热请求（供外部调功器）/ heating request for the power unit
    bCoolFanOn       : BOOL;                 // 降温风机请求 / cooling fan request
    bDoorOpenPermit  : BOOL;                 // 开门许可（温度已降到阈值以下）/ door open permit
    fRateNow         : REAL;                 // 当前升温速率 [°C/min] / current ramp rate [°C/min]
    bSeqDone         : BOOL;                 // 段序完成脉冲（单拍）/ sequence done pulse, single scan
    bError           : BOOL;                 // 故障标志（锁存类归并）/ fault flag
    uErrorId         : UDINT;                // 故障码，0 = 无故障 / error code, 0 = none
    eState           : E_DL_CuringState;     // 当前状态（供 HMI 诊断）/ current state
END_VAR
VAR
    fbTrigStart      : R_TRIG;               // 启动沿检测实例 / start edge detector
    fbTrigReset      : R_TRIG;               // 复位沿检测实例 / reset edge detector
    tonHold          : TON;                  // 保温计时实例 / dwell timer
    tonRateWin       : TON;                  // 速率评估窗（自复位 R188）/ rate evaluation window, self resetting
    eStateInt        : E_DL_CuringState;     // 主状态机内部当前态 / internal state
    fTempPrev        : REAL;                 // 上一拍温度快照 [°C] / previous temperature snapshot [°C]
    fDtMin           : REAL;                 // 采样周期折算 [min]，除子 / sample period in minutes, the divisor
    nSampleMs        : DINT;                 // 采样周期整毫秒 [ms] / sample period in milliseconds
    bTempBad         : BOOL;                 // 本拍温度非有限 / temperature non-finite this scan
    bRateOver        : BOOL;                 // 本拍速率超限 / ramp rate exceeded this scan
    bDoorViolation   : BOOL;                 // 本拍开门违规 / door interlock violation this scan
    bRateLatch       : BOOL;                 // 速率超限锁存内部副本 / internal rate latch
    bDoorLatch       : BOOL;                 // 开门违规锁存内部副本 / internal door latch
    bCfgBad          : BOOL;                 // 本拍组态非法 / config illegal this scan
    bCfgLatch        : BOOL;                 // 组态锁存（复位沿 + 组态改对解除）/ config latch
    bDoneT           : BOOL;                 // 完成脉冲内部副本（单拍）/ internal done pulse
    bErrorInt        : BOOL;                 // 本拍故障置位累加 / fault set accumulator
    bFirstScan       : BOOL := TRUE;         // 上电首扫标志 / first-scan flag
END_VAR
VAR CONSTANT
    DL_CO_FIN_LIM  : REAL := 1.0E30;         // REAL 幅值兜底判界 / REAL magnitude bound
    DL_CO_MS_PER_MIN : REAL := 60000.0;      // 毫秒每分钟折算常数 [ms/min] / milliseconds per minute
    DL_CO_RATE_EPS : REAL := 1.0E-6;         // 速率比较容差（浮点禁判等）/ rate comparison tolerance
END_VAR

(*------------------------------------------------------------------------------
 * 段 1｜无条件刷新区（红线 R7）：二沿二计时位于主体最前部
 *      Unconditional refresh: two edges and two timers at the very top
 *-----------------------------------------------------------------------------*)
fbTrigStart(CLK := bStartCmd);
fbTrigReset(CLK := bReset);
tonHold(IN := (eStateInt = E_DL_CuringState.eHold), PT := tHold);
tonRateWin(IN := NOT tonRateWin.Q, PT := tSample);    // 自复位速率评估窗（R188）/ self-resetting rate window

(* 段 2｜上电首扫 / first-scan init *)
IF bFirstScan THEN
    eStateInt  := E_DL_CuringState.eIdle;
    fTempPrev  := 0.0;
    fRateNow   := 0.0;
    bRateLatch := FALSE;
    bDoorLatch := FALSE;
    bFirstScan := FALSE;
END_IF

(* 段 3｜每拍预清（FB32-1）：单拍标志，禁入锁存 / per-scan preset *)
bErrorInt := FALSE;
bDoneT    := FALSE;

(*------------------------------------------------------------------------------
 * 段 4｜组态域闸（R151 全枚举）+ 解除路径（R152 自证可达）
 *      Config gate over every threshold and the sample period, with the clear path
 *-----------------------------------------------------------------------------*)
nSampleMs := TIME_TO_DINT(tSample);                       // TIME -> 整毫秒 [ms] / TIME to milliseconds
fDtMin    := DINT_TO_REAL(nSampleMs) / DL_CO_MS_PER_MIN;  // 毫秒 -> 分钟（除子常数 > 0）[min] / to minutes

bCfgBad := (fRateMax <= 0.0) OR (fRateMax <> fRateMax)
           OR (tHold <= T#0S)
           OR (fTempSet <> fTempSet) OR (ABS(fTempSet) >= DL_CO_FIN_LIM)
           OR (fDoorOpenTempMax <> fDoorOpenTempMax) OR (ABS(fDoorOpenTempMax) >= DL_CO_FIN_LIM)
           OR (tSample <= T#0S) OR (fDtMin <= 0.0) OR (fDtMin <> fDtMin);

IF bCfgBad THEN
    bCfgLatch := TRUE;
END_IF
IF fbTrigReset.Q AND (NOT bCfgBad) THEN
    bCfgLatch := FALSE;                    // 组态锁存解除 / config latch cleared
    uErrorId  := 16#0000_0000;             // 码位随解除归零 / code cleared with the latch
END_IF
IF bCfgLatch THEN
    uErrorId  := 16#0005_03B6;             // 故障级：组态非法 / fault: illegal configuration
    bErrorInt := TRUE;                     // R45 配对 / paired with the code
    eStateInt := E_DL_CuringState.eFault;
END_IF

(*------------------------------------------------------------------------------
 * 段 5｜判据求值：信号闸 + 速率 + 开门联锁（非有限只挂起不锁存）
 *      Criteria: signal gate, ramp rate and the door interlock
 *      速率只在评估窗到期拍折算一次（窗内保持不变），避免同拍差分放大噪声。
 *-----------------------------------------------------------------------------*)
bTempBad := (fTemp <> fTemp)
            OR ((fTemp - fTemp) <> (fTemp - fTemp))
            OR (ABS(fTemp) >= DL_CO_FIN_LIM);

IF (NOT bTempBad) AND tonRateWin.Q THEN
    fRateNow  := (fTemp - fTempPrev) / fDtMin;   // 差分折速率（除子已闸 > 0）[°C/min] / ramp rate
    fTempPrev := fTemp;                          // 快照推进（仅在有效样本上）/ snapshot advances on valid samples only
ELSIF bTempBad THEN
    uErrorId := 16#0005_04DF;                    // 信息级：温度非有限，判据挂起 / info: non-finite temperature
END_IF

bRateOver := (NOT bTempBad) AND (fRateNow > (fRateMax + DL_CO_RATE_EPS));
bDoorViolation := (NOT bTempBad) AND (NOT bDoorClosed)
                  AND (fTemp > (fDoorOpenTempMax + DL_CO_RATE_EPS));

(*------------------------------------------------------------------------------
 * 段 6｜主状态机（红线 R6）：ENUM + CASE + ELSE 兜底
 *      bStop 只迁相不清锁存（复位作用域声明见头注释披露 5）
 *-----------------------------------------------------------------------------*)
CASE eStateInt OF

    E_DL_CuringState.eIdle:
        IF bReset THEN
            bRateLatch := FALSE;                 // 空闲相复位允许清两类锁存 / idle reset clears both latches
            bDoorLatch := FALSE;
            uErrorId   := 16#0000_0000;
        END_IF
        IF bEnable AND (NOT bCfgLatch) AND (NOT bRateLatch) AND (NOT bDoorLatch)
           AND fbTrigStart.Q THEN
            fTempPrev := fTemp;                  // 启动拍取当前温度作速率基准 / seed the rate baseline
            eStateInt := E_DL_CuringState.eHeat;
        END_IF

    E_DL_CuringState.eHeat:
        IF bStopCmd OR (NOT bEnable) THEN
            eStateInt := E_DL_CuringState.eIdle;
        ELSIF fTemp >= fTempSet THEN
            eStateInt := E_DL_CuringState.eHold; // 达温进保温 / setpoint reached, dwell
        END_IF

    E_DL_CuringState.eHold:
        IF bStopCmd OR (NOT bEnable) THEN
            eStateInt := E_DL_CuringState.eIdle;
        ELSIF tonHold.Q THEN
            uErrorId  := 16#0005_04DE;           // 信息级：保温完成 / info: dwell finished
            eStateInt := E_DL_CuringState.eCool; // 进降温段 / to cooling
        END_IF

    E_DL_CuringState.eCool:
        IF bStopCmd OR (NOT bEnable) THEN
            eStateInt := E_DL_CuringState.eIdle;
        ELSIF fTemp <= fDoorOpenTempMax THEN
            eStateInt := E_DL_CuringState.eDone; // 温度达开门阈，段序完成 / cool enough, done
        END_IF

    E_DL_CuringState.eDone:
        bDoneT    := TRUE;                       // 完成脉冲：内部置位 -> 出口单拍（两段式）/ done pulse via the exit
        eStateInt := E_DL_CuringState.eIdle;     // 单拍完成相 / one-shot phase

    E_DL_CuringState.eFault:
        (* 解除路径（R152 自证可达）：复位沿 AND 组态改对 AND 两判据本拍均已消失 *)
        IF fbTrigReset.Q AND (NOT bCfgBad) AND (NOT bRateOver) AND (NOT bDoorViolation) THEN
            bCfgLatch  := FALSE;                 // 三类锁存同沿解除 / three latches cleared together
            bRateLatch := FALSE;
            bDoorLatch := FALSE;
            uErrorId   := 16#0000_0000;
            eStateInt  := E_DL_CuringState.eIdle;
        END_IF

    ELSE
        (* 非法状态拦截 / illegal state interception *)
        eStateInt := E_DL_CuringState.eFault;
        uErrorId  := 16#0005_03B6;
        bErrorInt := TRUE;

END_CASE;

(*------------------------------------------------------------------------------
 * 段 7｜锁存消化：速率超限与开门违规各自独立锁存 + 独立码位（R190 归因唯一）
 *      Latch digestion with two distinct causes and codes
 *-----------------------------------------------------------------------------*)
IF bRateOver AND (NOT bRateLatch) THEN
    bRateLatch := TRUE;                          // 速率超限锁存 / ramp rate latched
    uErrorId   := 16#0005_03B4;                  // 故障级：升温速率超限 / fault: ramp rate exceeded
    bErrorInt  := TRUE;                          // R45 配对 / paired with the code
    eStateInt  := E_DL_CuringState.eFault;
END_IF
IF bDoorViolation AND (NOT bDoorLatch) THEN
    bDoorLatch := TRUE;                          // 开门违规锁存 / door violation latched
    uErrorId   := 16#0005_03B5;                  // 故障级：降温未达标即开门 / fault: door opened too hot
    bErrorInt  := TRUE;                          // R45 配对 / paired with the code
    eStateInt  := E_DL_CuringState.eFault;
END_IF

(*------------------------------------------------------------------------------
 * 段 8｜输出单一出口（范式 P-05）：执行请求只由状态派生
 *      Single output exit: every request derives from the phase
 *-----------------------------------------------------------------------------*)
bHeatOn         := ((eStateInt = E_DL_CuringState.eHeat) OR (eStateInt = E_DL_CuringState.eHold))
                   AND (NOT bCfgLatch) AND (NOT bRateLatch);
bCoolFanOn      := (eStateInt = E_DL_CuringState.eCool) AND (NOT bCfgLatch);
bDoorOpenPermit := ((NOT bTempBad) AND (fTemp <= fDoorOpenTempMax))
                   AND (eStateInt <> E_DL_CuringState.eHeat) AND (eStateInt <> E_DL_CuringState.eHold)
                   AND (NOT bDoorLatch);
bSeqDone        := bDoneT;                       // 单拍脉冲统一出口 / unified single-scan exit
bError          := bErrorInt OR bCfgLatch OR bRateLatch OR bDoorLatch;
eState          := eStateInt;
END_FUNCTION_BLOCK

(* ---- FB_DL_CvdTempRamp.st ---- *)
(*
  FB_DL_CvdTempRamp  —  CVD/扩散炉多段 Ramp/Soak 曲线跟随 + 均匀性判据 / CVD furnace multi-segment ramp-soak tracking with uniformity
  分类 Category : DL_Process
  码位 Code     : 16#06_0_91
  版本 Version  : 1.0.0
  溯源 Source   : LGF Technology 语义借鉴 · clean-room 实现，仅借分类/参数域/命名，未复制源码
  功能 Function : 1) 多段 Ramp/Soak 工艺曲线跟随（复用 FB_DL_RampSoakProfile 设定源，全部温区共用同一条曲线）；
                  2) 均匀性判据：各温区统计均值与设定偏差逐区复核，全区进窗才置 bUniformOk；
                  3) Ramp 段跟随失败升级（|实测 − 设定| 持续超限 → 段故障锁存）。
  边界 Boundary : ① 均匀性测点 < 2 不出结论（信息级，禁单点冒充均匀性）；
                  ② 任一温区无效：该区判定冻结并置码，禁塞伪值；
                  ③ Ramp 段斜率跟随偏差超限持续 N 拍判跟随失败升级（非死等）；
                  ④ Soak 终点窗带独立超时出口（计时超限升级）；
                  ⑤ 与 FB_DL_LaminatorTempProfile 职责边界：本件面向 CVD/扩散炉多段（1..8 段可配）
                     工艺曲线 + 跨温区均匀性判据；层压机件为固定三段真空/加压配方 + 保温保持出口，
                     二者行业参数集与判据分立，互不替代。
  依赖 Depends  : FB_DL_RampSoakProfile × 1（设定源，每拍无条件调用）
                  FB_DL_SignalStatistics × 4（逐温区偏差统计，每拍无条件调用）

  码表 Error codes（本件子码步进 16#30 · 本格 91 与既有 9X 子码段冲突，错位至 C1/D1 避让）:
    16#0002_06C1 故障级：组态非法（段数越界 / 终点窗或跟随门限 <= 0 / 目标温度非有限）
    16#0002_06D1 故障级：跟随失败（Ramp 段偏差持续超门限）或 Soak 超时（锁存需复位）
    16#0002_06B1 信息级：温区无效判定冻结 / 有效测点 < 2 不出均匀性结论（不置 bError）
*)

TYPE E_DL_CtrPhase :
(
    eIdle   := 0,   // 空闲 / Idle
    eRun    := 10,  // 曲线跟随中 / Profile tracking
    eSoakOk := 20,  // 全区保温进窗 / All zones in soak window
    eDone   := 30,  // 曲线完成 / Profile done
    eFrozen := 40,  // 全部温区无效冻结 / All zones frozen
    eFault  := 90   // 跟随失败/超时锁定 / Tracking failure or timeout locked
);
END_TYPE

FUNCTION_BLOCK FB_DL_CvdTempRamp
VAR_INPUT
    bStart        : BOOL;                           // 启动指令，上升沿生效 / Profile start, edge
    bHold         : BOOL;                           // 外部保持 / External hold
    bReset        : BOOL;                           // 复位，上升沿清故障 / Reset, clears fault
    nSegCount     : INT := 4;                       // 有效段数 [段]，1..8 / Active segment count
    aSegTgtC      : ARRAY[1..8] OF REAL;            // 各段目标温度 [°C] / Segment targets [degC]
    aSegRampT     : ARRAY[1..8] OF TIME;            // 各段斜坡时间 [s]，0 = 阶跃直达 / Segment ramp times
    aSegSoakT     : ARRAY[1..8] OF TIME;            // 各段保温时间 [s]，0 = 无保温 / Segment soak times
    aZoneTempC    : ARRAY[1..4] OF REAL;            // 各温区实测温度 [°C] / Zone measured temperature [degC]
    nZoneCount    : INT := 4;                       // 温区数 [区]，1..4（均匀性测点数）/ Zone count
    fFollowMaxK   : REAL := 15.0;                   // Ramp 跟随偏差门限 [K]，域 > 0 / Tracking deviation limit [K]
    uFollowConfirm: UINT := 10;                     // 跟随失败确认拍数 [拍] / Tracking failure confirm scans
    fEndWinK      : REAL := 3.0;                    // Soak 终点窗半宽 [K]，域 > 0 / Soak end window half width [K]
    fEps          : REAL := 1.0E-6;                 // 浮点判零容差 [1] / Floating zero tolerance
END_VAR
VAR_OUTPUT
    fSetpointC    : REAL;                           // 曲线设定输出 [°C] / Profile setpoint output [degC]
    nSegAct       : INT;                            // 当前段号 1..nSegCount / Active segment
    bSoakInWindow : BOOL;                           // 全区保温进窗（多拍确认）/ All zones in soak window
    bUniformOk    : BOOL;                           // 均匀性结论（全区偏差窗内）/ Uniformity verdict
    bProfileDone  : BOOL;                           // 曲线完成标志（保持型）/ Profile done, held
    bError        : BOOL;                           // 故障标志，与故障级码配对 / Fault flag
    uErrorId      : UDINT;                          // 事件码，0 = 无事件 / Event code
    eStateOut     : E_DL_CtrPhase;                  // 状态机当前态，段尾单点映射 / Phase mapped at tail
END_VAR
VAR
    _eState       : E_DL_CtrPhase := E_DL_CtrPhase.eIdle;  // 内部状态 / Internal state
    fbRs          : FB_DL_RampSoakProfile;          // 曲线设定源实例（无条件调用）/ Profile setpoint source
    afbStat       : ARRAY[1..4] OF FB_DL_SignalStatistics;  // 逐温区偏差统计（无条件调用）/ Per-zone deviation statistics
    rtrStart      : R_TRIG;                         // 启动沿 / Start edge
    rtrReset      : R_TRIG;                         // 复位沿 / Reset edge
    abZoneOk      : ARRAY[1..4] OF BOOL;            // 温区有效掩码 / Zone validity mask
    abZoneInWin   : ARRAY[1..4] OF BOOL;            // 温区进窗掩码 / Zone in-window mask
    bCfgOk        : BOOL;                           // 组态合法标志 / Configuration valid
    bAnyOk        : BOOL;                           // 存在有效温区 / Any valid zone
    bAllInvalid   : BOOL;                           // 全部温区无效 / All zones invalid
    bInRamp       : BOOL;                           // 本拍处于 Ramp 段 / In ramp segment this scan
    bDevOver      : BOOL;                           // 跟随偏差超限（电平）/ Deviation over limit
    uFollowCnt    : UINT;                           // 跟随失败确认计数 [拍] / Tracking failure counter
    bSoakTout     : BOOL;                           // Soak 终点窗超时 / Soak end-window timeout
    fSoakElapsed  : REAL;                           // 进窗后累计等待 [s] / Elapsed wait after in-window [s]
    nZ            : INT;                            // 温区遍历索引 / Zone loop index
    uFault        : UDINT;                          // 锁存故障码 / Latched fault code
    uInfo         : UDINT;                          // 信息级码 / Information code
END_VAR
VAR CONSTANT
    DL_CTR_ZMAX   : INT := 4;                       // 温区数上限 [区] / Zone count upper bound
    DL_CTR_INFMAX : REAL := 1.0E30;                 // 温度有限值幅值上限 [°C] / Temperature finite bound [degC]
    DL_CTR_SOAK_TOUT : REAL := 60.0;                // Soak 终点窗独立超时 [s] / Soak end-window timeout [s]
END_VAR

(* === 段 0 · 实例刷新 === *)
rtrStart(CLK := bStart);                          // 每拍刷新启动沿
rtrReset(CLK := bReset);                          // 每拍刷新复位沿

(* === 段 1 · 组态闸 === *)
bCfgOk := (nSegCount >= 1) AND (nSegCount <= 8)   // 段数域闸
          AND (nZoneCount >= 1) AND (nZoneCount <= DL_CTR_ZMAX)
          AND (fFollowMaxK > fEps) AND (fEndWinK > fEps)       // 门限正域
          AND (fbRs.fSetpoint = fbRs.fSetpoint);  // 实例侧哨兵（首拍未运行恒真）
FOR nZ := 1 TO 8 DO
    bCfgOk := bCfgOk AND (aSegTgtC[nZ] = aSegTgtC[nZ])         // 段目标 NaN 自反
              AND (ABS(aSegTgtC[nZ]) < DL_CTR_INFMAX);         // 段目标幅值域
END_FOR
IF NOT bCfgOk THEN
    uFault := 16#0002_06C1;                       // 故障级：组态非法
END_IF
IF rtrReset.Q AND bCfgOk THEN
    uFault := 16#0000;                            // 复位沿清锁存（解除路径可达）
    uFollowCnt := UINT#0;                         // 跟随确认计数复位
    fSoakElapsed := 0.0;                          // 进窗等待清零
    FOR nZ := 1 TO DL_CTR_ZMAX DO
        abZoneInWin[nZ] := FALSE;                 // 进窗掩码复位
    END_FOR
END_IF
uInfo := 16#0000;                                 // 信息码每拍清零

(* === 段 2 · 曲线设定源实例（无条件调用）与温区域闸 === *)
fbRs(bStart := rtrStart.Q,                        // 启动沿透传
     bHold := bHold,                              // 外部保持透传
     fStartValue := aZoneTempC[1],                // 首段斜坡起点取 1 区实测（无效时实例域闸兜底）
     nSegCount := INT_TO_USINT(MAX(nSegCount, 1)),// 段数下限防 0
     aTarget := aSegTgtC,                         // 段目标表
     aRampTime := aSegRampT,                      // 段斜坡表
     aSoakTime := aSegSoakT,                      // 段保温表
     bLoopProfile := FALSE,                       // 单次工艺曲线不循环
     bReset := rtrReset.Q);                       // 复位沿透传
fSetpointC := fbRs.fSetpoint;                     // 设定输出
nSegAct := fbRs.nSegAct;                          // 段号输出
bInRamp := (fbRs.ePhase = E_DL_RampSoakPhase.eRamp);  // Ramp 相判据（枚举成员对齐属主件）
bAnyOk := FALSE;                                  // 有效区汇总先清
bAllInvalid := TRUE;                              // 全无效假设先置
FOR nZ := 1 TO DL_CTR_ZMAX DO
    abZoneOk[nZ] := (nZ <= nZoneCount)
                    AND (aZoneTempC[nZ] = aZoneTempC[nZ])
                    AND (ABS(aZoneTempC[nZ]) < DL_CTR_INFMAX);  // NaN 自反 + 幅值闸
    bAnyOk := bAnyOk OR abZoneOk[nZ];             // 汇总有效
    bAllInvalid := bAllInvalid AND (NOT abZoneOk[nZ]);  // 汇总全无效
    afbStat[nZ](fIn := aZoneTempC[nZ] - fSetpointC,             // 偏差量统计（无效值由实例域闸拒绝）
                bSample := abZoneOk[nZ] AND (NOT bHold),        // 无效/保持拍不采
                nWindow := 16,                    // 偏差窗 16 样本
                bClear := rtrStart.Q);            // 启动沿清窗重计
    abZoneInWin[nZ] := abZoneOk[nZ] AND afbStat[nZ].bValid
                       AND (ABS(afbStat[nZ].fMean) <= fEndWinK + fEps);  // 均值偏差进窗
END_FOR
IF bAllInvalid THEN
    uInfo := 16#0002_06B1;                        // 信息级：温区无效判定冻结
END_IF

(* === 段 3 · 全区进窗汇总 / 跟随失败与 Soak 超时判据 === *)
bSoakInWindow := (nZoneCount >= 2) AND (NOT bAllInvalid);      // 测点 < 2 不出进窗结论
FOR nZ := 1 TO nZoneCount DO
    bSoakInWindow := bSoakInWindow AND abZoneInWin[nZ];        // 全区进窗才成立
END_FOR
IF (NOT bSoakInWindow) AND (nZoneCount < 2) AND bAnyOk THEN
    uInfo := 16#0002_06B1;                        // 信息级：有效测点不足不出结论
END_IF
bDevOver := FALSE;                                // 跟随偏差超限本拍重算
FOR nZ := 1 TO nZoneCount DO
    bDevOver := bDevOver OR (abZoneOk[nZ] AND afbStat[nZ].bValid
               AND (ABS(afbStat[nZ].fMean) > fFollowMaxK));      // 任一有效区均值偏差超门限
END_FOR
IF bInRamp AND bDevOver THEN
    uFollowCnt := uFollowCnt + UINT#1;            // Ramp 段偏差超限确认计数
    IF uFollowCnt >= uFollowConfirm THEN
        uFault := 16#0002_06D1;                   // 故障级：跟随失败升级（锁存，非死等）
    END_IF
ELSE
    uFollowCnt := UINT#0;                         // 未超限/非 Ramp 段：计数归零
END_IF
bSoakTout := FALSE;                               // Soak 超时本拍重算
IF bSoakInWindow THEN
    fSoakElapsed := fSoakElapsed + 0.1;           // 进窗后等待累计（周期 0.1 s 口径，与实例采样对齐）
    IF fSoakElapsed > DL_CTR_SOAK_TOUT THEN
        bSoakTout := TRUE;                        // 终点窗独立超时出口
        uFault := 16#0002_06D1;                   // 故障级：Soak 超时（锁存）
    END_IF
ELSE
    fSoakElapsed := 0.0;                          // 未持续进窗：等待清零
END_IF

(* === 段 4 · 主状态机（ENUM + CASE，含 ELSE 兜底）=== *)
CASE _eState OF
E_DL_CtrPhase.eIdle :
    bProfileDone := FALSE;                        // 空闲未完成
    bSoakInWindow := FALSE;                       // 空闲无进窗
    IF uFault <> 16#0000 THEN
        _eState := E_DL_CtrPhase.eFault;          // 故障优先
    ELSIF fbRs.nSegAct > 0 THEN
        _eState := E_DL_CtrPhase.eRun;            // 设定源已启动进运行相
    END_IF

E_DL_CtrPhase.eRun :
    bUniformOk := bSoakInWindow;                  // 均匀性结论与进窗同判据（均值偏差窗）
    IF uFault <> 16#0000 THEN
        _eState := E_DL_CtrPhase.eFault;          // 跟随失败/超时转故障
    ELSIF bAllInvalid THEN
        _eState := E_DL_CtrPhase.eFrozen;         // 全区无效转冻结
    ELSIF fbRs.bDone THEN
        bProfileDone := TRUE;                     // 曲线完成（保持型）
        _eState := E_DL_CtrPhase.eDone;           // 转完成相
    ELSIF bSoakInWindow THEN
        _eState := E_DL_CtrPhase.eSoakOk;         // 全区进窗转保温合格相
    END_IF

E_DL_CtrPhase.eSoakOk :
    bUniformOk := TRUE;                           // 均匀性保持
    bSoakInWindow := TRUE;                        // 进窗保持（防同拍抹除）
    IF uFault <> 16#0000 THEN
        _eState := E_DL_CtrPhase.eFault;          // 故障转出
    ELSIF fbRs.bDone THEN
        bProfileDone := TRUE;                     // 曲线完成
        _eState := E_DL_CtrPhase.eDone;           // 转完成相
    ELSIF NOT bAnyOk THEN
        _eState := E_DL_CtrPhase.eFrozen;         // 全区无效转冻结
    END_IF

E_DL_CtrPhase.eDone :
    bProfileDone := TRUE;                         // 完成保持
    IF rtrStart.Q THEN
        bProfileDone := FALSE;                    // 新启动沿重开
        _eState := E_DL_CtrPhase.eRun;            // 回运行相
    END_IF

E_DL_CtrPhase.eFrozen :
    bProfileDone := FALSE;                        // 冻结相不出完成
    bSoakInWindow := FALSE;                       // 冻结相不出进窗
    IF bAnyOk AND (uFault = 16#0000) THEN
        _eState := E_DL_CtrPhase.eRun;            // 任一区恢复回运行（解除路径可达）
    END_IF

E_DL_CtrPhase.eFault :
    bSoakInWindow := FALSE;                       // 故障相不出进窗
    IF uFault = 16#0000 THEN
        _eState := E_DL_CtrPhase.eIdle;           // 解锁回空闲
    END_IF

ELSE
    _eState := E_DL_CtrPhase.eFault;              // 非法状态拦截
    uFault := 16#0002_06C1;                       // 故障级：相 ID 越界复用组态码段
END_CASE

(* === 段 5 · 输出映射 === *)
bError := (uFault <> 16#0000);                    // 故障标志仅由故障级码置位（R45 配对）
IF bError THEN
    uErrorId := uFault;                           // 故障级优先上报
ELSE
    uErrorId := uInfo;                            // 否则上报信息级码
END_IF
eStateOut := _eState;                             // 输出枚举段尾单点映射（N2 规则）
END_FUNCTION_BLOCK
